Universal Robots URScript: test.script

def test():
  global _hidden_verificationVariable=0
  step_count_363709d2_59a1_48ba_b260_6a0887d41453 = 0.0
  thread Step_Counter_Thread_5b3f90a0_63de_4def_b0b2_14eef1768a44():
    while (True):
      step_count_363709d2_59a1_48ba_b260_6a0887d41453 = step_count_363709d2_59a1_48ba_b260_6a0887d41453 + 1.0
      sync()
    end
  end
  run Step_Counter_Thread_5b3f90a0_63de_4def_b0b2_14eef1768a44()
  set_gravity([0.0, 0.0, 9.82])
  motion_version_set(1)
  tool_wrench_limit_disable()
  set_tcp(p[0.0,0.0,0.161,3.1415,0.0,0.0])
  set_safety_mode_transition_hardness(1)
  set_standard_analog_input_domain(0, 1)
  set_standard_analog_input_domain(1, 1)
  set_tool_analog_input_domain(0, 1)
  set_tool_analog_input_domain(1, 1)
  set_analog_outputdomain(0, 1)
  set_analog_outputdomain(1, 1)
  set_input_actions_to_default()
  set_standard_digital_input_action(0, "freedrive")
  set_gp_boolean_input_action(0, "freedrive")
  set_runstate_standard_digital_outputs([0])
  set_runstate_configurable_digital_outputs([5])
  set_runstate_standard_digital_output_to_value(0, 1)
  set_runstate_configurable_digital_output_to_value(5, 1)
  set_runstate_configurable_digital_output_to_value(6, 2)
  set_runstate_configurable_digital_output_to_value(7, 2)
  modbus_add_signal("192.168.12.20", 255, 3, 2, "MiR_Mode", False)
  modbus_set_signal_update_frequency("MiR_Mode", 10)
  modbus_add_signal("192.168.12.20", 255, 4, 2, "MiR_State", False)
  modbus_set_signal_update_frequency("MiR_State", 10)
  modbus_add_signal("192.168.12.20", 255, 5, 2, "MiR_Error_ID", False)
  modbus_set_signal_update_frequency("MiR_Error_ID", 10)
  modbus_add_signal("192.168.12.20", 255, 7, 2, "MiR_Battery_Lvl", False)
  modbus_set_signal_update_frequency("MiR_Battery_Lvl", 10)
  modbus_add_signal("192.168.12.20", 255, 18, 2, "MiR_Mis_Queue", False)
  modbus_set_signal_update_frequency("MiR_Mis_Queue", 10)
  modbus_add_signal("192.168.12.20", 255, 1, 1, "MiR_CMD_Stop", False)
  modbus_set_signal_update_frequency("MiR_CMD_Stop", 10)
  modbus_add_signal("192.168.12.20", 255, 2, 1, "MiR_CMD_Abort", False)
  modbus_set_signal_update_frequency("MiR_CMD_Abort", 10)
  modbus_add_signal("192.168.12.20", 255, 3, 1, "MiR_CMD_Clear_Q", False)
  modbus_set_signal_update_frequency("MiR_CMD_Clear_Q", 10)
  modbus_add_signal("192.168.12.20", 255, 4, 1, "MiR_CMD_Clear_E", False)
  modbus_set_signal_update_frequency("MiR_CMD_Clear_E", 10)
  modbus_add_signal("192.168.12.20", 255, 5, 1, "MiR_CMD_Start", False)
  modbus_set_signal_update_frequency("MiR_CMD_Start", 10)
  modbus_add_signal("192.168.12.20", 255, 1001, 2, "T2O_Current_Pos", False)
  modbus_set_signal_update_frequency("T2O_Current_Pos", 10)
  modbus_add_signal("192.168.12.20", 255, 1003, 2, "T2O_Warning_ID", False)
  modbus_set_signal_update_frequency("T2O_Warning_ID", 10)
  modbus_add_signal("192.168.12.20", 255, 1005, 2, "T2O_Error_ID", False)
  modbus_set_signal_update_frequency("T2O_Error_ID", 10)
  modbus_add_signal("192.168.12.20", 255, 1019, 3, "O2T_Target_Pos", False)
  modbus_set_signal_update_frequency("O2T_Target_Pos", 10)
  modbus_add_signal("192.168.12.20", 255, 1017, 3, "O2T_Action", False)
  modbus_set_signal_update_frequency("O2T_Action", 10)
  modbus_add_signal("192.168.12.20", 255, 1000, 1, "O2T_Mis_Charge", False)
  modbus_set_signal_update_frequency("O2T_Mis_Charge", 1)
  modbus_add_signal("192.168.12.20", 255, 1004, 1, "O2T_Mis_Main", False)
  modbus_set_signal_update_frequency("O2T_Mis_Main", 1)
  modbus_add_signal("192.168.12.20", 255, 1007, 2, "T2O_Nav_Attemps", False)
  modbus_set_signal_update_frequency("T2O_Nav_Attemps", 10)
  modbus_add_signal("192.168.12.20", 255, 1009, 2, "T2O_Done", False)
  modbus_set_signal_update_frequency("T2O_Done", 10)
  modbus_add_signal("192.168.12.20", 255, 1021, 3, "O2T_Acknowledge", False)
  modbus_set_signal_update_frequency("O2T_Acknowledge", 10)
  modbus_add_signal("192.168.12.20", 255, 1011, 2, "T2O_Charging", False)
  modbus_set_signal_update_frequency("T2O_Charging", 10)
  modbus_add_signal("192.168.12.20", 255, 12, 2, "MiR_Position_X1", False)
  modbus_set_signal_update_frequency("MiR_Position_X1", 10)
  modbus_add_signal("192.168.12.20", 255, 13, 2, "MiR_Position_X2", False)
  modbus_set_signal_update_frequency("MiR_Position_X2", 10)
  modbus_add_signal("192.168.12.20", 255, 14, 2, "MiR_Position_Y1", False)
  modbus_set_signal_update_frequency("MiR_Position_Y1", 10)
  modbus_add_signal("192.168.12.20", 255, 15, 2, "MiR_Position_Y2", False)
  modbus_set_signal_update_frequency("MiR_Position_Y2", 10)
  modbus_add_signal("192.168.12.20", 255, 1023, 3, "O2T_Footprint", False)
  modbus_set_signal_update_frequency("O2T_Footprint", 10)
  modbus_add_signal("192.168.12.20", 255, 1025, 3, "O2T_ProtectOff", False)
  modbus_set_signal_update_frequency("O2T_ProtectOff", 10)
  modbus_add_signal("192.168.12.20", 255, 1027, 3, "O2T_Dock", False)
  modbus_set_signal_update_frequency("O2T_Dock", 10)
  modbus_add_signal("192.168.12.20", 255, 16, 2, "MiR_Theta_1", False)
  modbus_set_signal_update_frequency("MiR_Theta_1", 10)
  modbus_add_signal("192.168.12.20", 255, 17, 2, "MiR_Theta_2", False)
  modbus_set_signal_update_frequency("MiR_Theta_2", 10)
  modbus_add_signal("192.168.12.197", 255, 0, 0, "WM_Sensor1", False)
  modbus_set_signal_update_frequency("WM_Sensor1", 2)
  modbus_add_signal("192.168.12.197", 255, 1, 0, "WM_Sensor2", False)
  modbus_set_signal_update_frequency("WM_Sensor2", 2)
  modbus_add_signal("192.168.12.197", 255, 2, 0, "WM_Sensor3", False)
  modbus_set_signal_update_frequency("WM_Sensor3", 2)
  modbus_set_runstate_dependent_choice("MiR_CMD_Stop",0)
  modbus_set_runstate_dependent_choice("MiR_CMD_Abort",0)
  modbus_set_runstate_dependent_choice("MiR_CMD_Clear_Q",0)
  modbus_set_runstate_dependent_choice("MiR_CMD_Clear_E",0)
  modbus_set_runstate_dependent_choice("MiR_CMD_Start",0)
  modbus_set_runstate_dependent_choice("O2T_Target_Pos",0)
  modbus_set_runstate_dependent_choice("O2T_Action",0)
  modbus_set_runstate_dependent_choice("O2T_Mis_Charge",0)
  modbus_set_runstate_dependent_choice("O2T_Mis_Main",0)
  modbus_set_runstate_dependent_choice("O2T_Acknowledge",0)
  modbus_set_runstate_dependent_choice("O2T_Footprint",0)
  modbus_set_runstate_dependent_choice("O2T_ProtectOff",0)
  modbus_set_runstate_dependent_choice("O2T_Dock",0)
  set_target_payload(1.480000, [-0.002000, 0.016000, 0.051000], [0.002959, 0.002959, 0.002959, 0.000000, 0.000000, 0.000000])
  set_tool_communication(True, 115200, 0, 1, 1.5, 3.5)
  set_tool_output_mode(0)
  set_tool_digital_output_mode(0, 1)
  set_tool_digital_output_mode(1, 1)
  set_tool_voltage(24)
  global AMR_AtTarget=False
  global ARM_Referenced=False
  global PROCESS_Info=""
  global AMR_Step=0
  global STATE=4
  global AMR_Free=False
  global AMR_PosTarget=0
  global PSE_G_H=p[0, 0, 0, 0, 0, 0]
  global PSE_T=p[0.00001, -0.4, 0.30003, -0.00005, 0.00001, 0.00002]
  global PSE_R=p[0, 0, 0, 0, 0, 0]
  global AMR_PosActual=7
  global PSE_G=p[0, 0, 0, 0, 0, 0]
  global PSE_A=p[0, 0, 0, 0, 0, 0]
  global PSE_C_S=p[0, 0, 0, 0, 0, 0]
  global PSE_C_H=p[0, 0, 0, 0, 0, 0]
  global PSE_C_E=p[0, 0, 0, 0, 0, 0]
  global PSE_T_H=p[0, 0, 0, 0, 0, 0]
  global AMR_Done=True
  global STATE_Info="Idle"
  global PROCESS_Step=0
  global PSE_A_H=p[0, 0, 0, 0, 0, 0]
  global PSE_R_H=p[0, 0, 0, 0, 0, 0]
  global JNT_A=[0, 0, 0, 0, 0, 0]
  global JNT_S=[0, 0, 0, 0, 0, 0]
  global ITM_ID=0
  global JIG=0
  global JIG_Slot=0
  global OBJ_Type=0
  global PSE_Z=p[0, 0, 0, 0, 0, 0]
  global CAM_LM_Detected=True
  global CAM_LM_ID=0
  global CAM_LM_Refinmnt=False
  global CAM_Captures=0
  global CAM_Done=True
  global CAM_LM_Refined=False
  global CAM_PRM_Retries=15
  global AMR_Battery=100
  global WRK_Done=False
  global ITM_Prepared=False
  global ITM_Manipulated=False
  global AMR_Charging=False
  global Action=0
  global Task_info=""
  global Action_Info=""
  global OBJ_Picked=False
  global TM_St_Stopping="0/2/50/2"
  global STATE_Times=[37070.92578, 339840.90625, 1824.11072, 1448747.625, 26510.78125, 599104.5625, 7693.4209, 27714.24023, 201.30833, 28483.10742, 31.506, 0.258, 385.68799, 0.256, 0, 0, 0]
  global TM_St_Stopped="3/22/24/0"
  global TM_St_Resetting="0/0/30/24"
  global TM_St_Idle="16/18/25/47"
  global TM_St_Starting="0/7/21/50"
  global TM_St_Execute="6/22/25/4"
  global TM_St_Holding="0/0/3/21"
  global TM_St_Held="0/7/54/43"
  global TM_St_Unholding="0/0/0/31"
  global TM_St_Suspendin="0/0/0/0"
  global TM_St_Suspended="0/0/6/25"
  global TM_St_Unsuspend="0/0/0/0"
  global TM_St_Completin="0/2/8/13"
  global TM_St_Complete="0/7/41/54"
  global TM_St_Aborting="00/00/00/00"
  global TM_St_Aborted="00/00/00/00"
  global TM_St_Clearing="00/00/00/00"
  global CMD_Stop=False
  global STP_Info=""
  global WRK_Step=0
  global WRK_Info=""
  global AMR_FootprintID=1
  global JNT_Z=[0, 0, 0, 0, 0, 0]
  global CAM_LM_Offset=p[0, 0, 0, 0, 0, 0]
  global CAM_LM_Deviatn=p[0, 0, 0, 0, 0, 0]
  global ITM_ID_List=[1, 2, 3, 4, 5, 6, 7, 8, 9]
  global JNT_Q=[0, 0, 0, 0, 0, 0]
  global OBJ_TCP=p[0, 0.08604, 0.29117, 0, -3.14159, 0]
  global OBJ_GRP_Offset=p[0, 0, 0.15, 0, 0, 0]
  global Task_ID=0
  global PRC_Force_Decap=False
  global PRC_Reset=True
  global CAM_CNT_Obj=0
  global OBJ_Nbr=0
  global GRP_Offset=p[0, 0, 0, 0, 0, 0]
  global GRP_Open_Pos=6
  global CMD_Hold=False
  global CAM_OBJ_Color="135639"
  global JIG_Offset=p[0, 0, 0, 0, 0, 0]
  global PRM_TO_Read_BC=5
  global OBJ_Brc_OK=True
  global SERVER_IP="192.168.12.139"
  global SERVER_PORT=3002
  global POTS_IP="192.168.12.102"
  global POTS_PORT=80
  global CAM_LM_SSRack=p[0.0,0.0,0.0,0.0,0.0,0.0]
  global Cont_A_TCP=p[-0.01446224178958122,-0.6317070151410098,0.23000037816712549,-1.0906492400659007,1.4047772946314183,-1.4136947877620298]
  global Cont_B_TCP=p[0.1998,-0.5012300000000001,0.21554327201208615,-1.2092122839110917,1.2091442884557517,-1.2093098736837602]
  global Cont_C_TCP=p[0.20899409891862653,-0.36521718091627275,0.22999234057600015,-1.2337601399754432,1.1952721569824734,-1.2073910748355074]
  global Decap_TCP_align=p[-0.041471808940011026,-0.3381541550735332,0.26582523339977177,-0.8796833786644639,1.6463420679311218,-1.709080917063812]
  global FRM_Cap_SSRack=p[0.5539194080315334,0.31767425178306713,0.33208398177541654,4.365192798093082E-5,-2.191282886828362E-5,0.8765357336623923]
  global FRM_Capture_Cen=p[-0.350002433865069,0.09999194422544704,0.39999652960929194,0.27390617458472216,0.27390634457500074,1.5534190527760867]
  global FRM_Capture_IN=p[0.14713742172916425,-0.4519990092180261,0.4999842175595519,1.716719843449274E-5,-5.967839199117233E-5,-3.141512274892885]
  global FRM_Centrifuge=p[-0.7614196357228254,0.13174165134832883,-0.40322998589848,0.051405105423226086,-0.012254257775454075,1.5210337802987177]
  global FRM_Container=p[-0.5003348223692186,0.35061804815168285,0.41579001388808423,-5.092943187272062E-5,1.0145185065363121E-4,-2.764319258713288]
  global FRM_Container_b=p[-0.5003368531143569,0.35061894438330765,0.41578806736276164,-8.54682865507139E-5,1.0209605772896093E-4,-2.8884715402158117]
  global FRM_PoTS=p[-0.5403054403210852,-0.10910773999775857,0.4828,3.058497512721046E-6,2.3454853329357316E-5,-2.208510541952706]
  global FRM_Reference=p[0.0,0.0,0.0,0.0,5.936340598853489E-5,0.0]
  global FRM_SS_SSTable=p[0.20318441097787696,-0.4018484849551291,0.0986494053372641,3.321622010808724E-5,1.2630310370280906E-5,2.9057826587464487E-5]
  global FRM_SWAB=p[-0.5425658438438228,0.050215382883637555,0.4828117991467299,1.2014498510989115E-5,1.8611655946156755E-5,-2.2084947047695405]
  global FRM_weigh_scale=p[-0.3804866881697204,0.025744252835212,0.4723487455232425,-1.0445769542396123E-4,-1.924788411074358E-5,-2.1691978730572363]
  global Home_Center=p[8.153119343667444E-6,-0.39999432384352546,0.2999959692487133,2.5646064776662724E-5,4.3940218780729606E-7,1.0264337438974612E-5]
  global Position1=p[-0.013283381383284571,-0.5604926192866768,0.38388715699602394,4.2328981461085945E-5,2.7078270325215812E-5,-3.7205146207707955E-5]
  global Position2=p[0.20351564705697425,-0.4203376101670667,0.3838762041571461,3.798288302544451E-5,4.704460451857417E-5,4.231147149799096E-6]
  global Position3=p[0.20350843333470736,-0.29021893349684563,0.38387753498709576,1.6019315164720892E-6,5.362200339537394E-5,1.3194338684148116E-5]
  global SAF_ULM_Back=p[0.0,0.25,0.0,-1.5707963267948966,0.0,0.0]
  global SAF_ULM_Bottom=p[0.0,0.0,0.175,0.0,-3.1411853059779946,6.144646783253781E-5]
  global SAF_ULM_Front=p[0.0,-0.8,0.0,1.5707963267948966,0.0,0.0]
  global SAF_ULM_Left=p[0.4,0.0,0.0,0.0,1.5707963267948966,0.0]
  global SAF_ULM_Right=p[-0.4,0.0,0.0,0.0,-1.5707963267948966,0.0]
  global Swab_Hol_NewApp=p[0.24367285099070987,-0.39538254967913455,0.1791890228280021,9.694511507909782E-6,-1.918651308171816E-5,-8.936699871509937E-5]
  global Swab_Holder=p[0.24295783117309838,-0.3013564682530984,0.1852322720229175,2.781519887568103E-5,4.9787017742599154E-5,-4.37903285531786E-5]
  global Swab_Holder_App=p[0.2429619714479549,-0.37982819606840945,0.18525382710668278,1.9222871262119376E-5,1.6223417670491008E-5,-5.4734062838048446E-5]
  global Swab_New_FlipAp=p[0.2397112683246373,-0.4131931547204771,0.1791901367353106,-3.2195134883720305E-6,5.5826332611522435E-5,3.121155597546625]
  global Swab_New_FlipHL=p[0.24201994270482732,-0.3016396679914842,0.1792041435801504,-5.840580747813655E-5,7.149594627182296E-5,3.1212173415187716]
  global Swab_flip_app=p[0.2429388733172488,-0.30137068448833126,0.2604132558601291,2.6401756342031075E-4,-5.484374510519208E-5,3.1254804120366084]
  global Swab_flip_hold=p[0.24294214110481466,-0.30136164018491357,0.18562266741928893,2.522236506414148E-4,-7.112060556159522E-5,3.1255321079816243]
  global Swab_holder_New=p[0.24365536646762584,-0.2997701233168029,0.17918094816818864,3.214234787213423E-5,4.175157661863989E-5,-5.646064180042735E-5]
  global Swab_take=p[0.06323186369735694,-0.63186492852859,0.1186768659332022,-0.0941457732311389,0.09836792894816203,-1.517326737506051]
  global Swab_take_appro=p[0.06320391400111934,-0.6318588436631464,0.19565149002631285,-0.09417297851843164,0.09839511960035544,-1.5173200644593776]
  global Trigger=p[0.0,0.0,0.0,0.0,0.0,0.0]
  global ULM_3FG=p[-0.030765235416747628,-0.34863465891472667,0.113,7.284395488044268E-6,3.273453749838684E-5,-1.4353257859996407]
  global ULM_Cap_Bin=p[-0.09250864937066318,-0.4278810928466919,0.11,0.012411963638116327,0.0011373915061224443,2.7934337459497622]
  global ULM_Cent_Racks=p[-0.18545280836253272,-0.6127182427471424,0.0092,-2.5489681018192384E-4,1.5011949774034494E-5,0.002017828229688311]
  global ULM_Input=p[0.24211961776286645,-0.49122804302630946,0.069,-0.0024427818584600467,0.009435707692609437,1.553764323389261]
  global ULM_NoK=p[-0.13173558762545426,-0.4223773499069831,0.1783860505865236,-0.013295546620598609,-0.0036702711105456223,-3.139406935149283]
  global ULM_Output=p[-0.03848915736486644,-0.4320501686344275,0.0,-6.433221303631731E-5,4.4743073056790854E-4,-3.1218466433891914]
  global ULM_SS_Jig=p[0.20042235181396445,-0.401422571467659,0.10172961048670293,-0.004383916608756479,-0.025399236865877438,0.14513627174952076]
  global swab_brk1=p[-0.038192766284940796,-0.35032292650225555,0.1065863357332553,-1.0289939058230132E-4,2.813749403516853,1.8382182448234926E-4]
  global uLM_Cap_SSRack=p[0.20881778585250285,-0.4048217020440386,0.5540171693698591,2.8523205665698764E-5,1.4454354491120644E-5,-0.034379521481452686]
  global uLM_SS_PickPlc=p[0.16950832747543634,-0.42825836359263725,0.10175705391961387,4.604858547296167E-4,-6.723821859499963E-4,-2.834490280150995]
  # begin: URCap Installation Node
  #   Source: UR Connect, 2.3.3, Universal Robots
  #   Type: UR Connect
  myurRPC = rpc_factory("xmlrpc","http://127.0.0.1:40474")
  # end: URCap Installation Node
  # begin: URCap Installation Node
  #   Source: Robotiq_Grippers, 3.17.0.105337, Robotiq Inc.
  #   Type: Vacuum
  #################################################
  # Vacuum Grip Check
  #################################################

  vacuumGripCheckThread1 = 0
  vacuumGripCheckThread2 = 0
  vacuumGripCheckThread3 = 0
  vacuumGripCheckThread4 = 0
  vacuumGripCheckThread1Running = False
  vacuumGripCheckThread2Running = False
  vacuumGripCheckThread3Running = False
  vacuumGripCheckThread4Running = False
  vacuumGripCheckSocketId = "1"
  vacuumGripCheckThreadStarted = False

  thread vacuumGripCheck():
    gripper_socket = vacuumGripCheckSocketId
    vacuumGripCheckThreadStarted = True

    while (True):
      objectDetectedDebounceCtr = 0

      while (objectDetectedDebounceCtr < 3):
        if(rq_is_vacuum_obj_detected(gripper_socket="1")):
          objectDetectedDebounceCtr = objectDetectedDebounceCtr + 1
        else:
          objectDetectedDebounceCtr = 0
        end
        sleep(0.1)
      end

      objectNotDetectedDebounceCtr = 0

      while objectNotDetectedDebounceCtr < 3:
        if (not rq_is_vacuum_obj_detected(gripper_socket="1")):
          objectNotDetectedDebounceCtr = objectNotDetectedDebounceCtr + 1
        else:
          objectNotDetectedDebounceCtr = 0
        end
        sleep(0.1)
      end

      socket_open("127.0.0.1",29999,"dashboardServerSocket")
      socket_send_line("pause","dashboardServerSocket")
      socket_send_string("popup Vacuum grip check has detected an object drop.", "dashboardServerSocket")
      socket_send_byte(10, "dashboardServerSocket")
      socket_close("dashboardServerSocket")

      sleep(0.008)
    end
  end

  def startVacuumGripCheckThread(gripperId="1"):
    vacuumGripCheckSocketId = gripperId
    threadHandle = run vacuumGripCheck()
    waitForVacuumGripCheckThreadStarted()
    return threadHandle
  end

  def stopVacuumGripCheckThread(threadHandle):
    kill threadHandle
  end

  def waitForVacuumGripCheckThreadStarted():
    while (not(vacuumGripCheckThreadStarted)):
      sleep(0.008)
    end
    vacuumGripCheckThreadStarted = False
  end
  #################################################
  # End - Vacuum Grip Check
  #################################################

  #################################################
  # Stops the pump on a distance travelled
  #################################################
  global stopPumpDistance = 100
  global stopPumpSocketId = "0"
  global stopPumpThreadStarted = [False, False, False, False]
  global stopPumpThreadHandles = [0, 0, 0, 0]

  thread stopPumpOnDistanceTravelled():
    distance = stopPumpDistance
    socketId = stopPumpSocketId
    stopPumpThreadStarted[rq_socket_to_index(socketId)] = True

    measuredDistance = waitForDistanceTravelled(distance)

    rq_stop(socketId)

    stopPumpThreadStarted[rq_socket_to_index(socketId)] = False
  end

  def waitForDistanceTravelled(distance):
    startingPose = get_actual_tcp_pose()
    measuredDistance = 0
    while (measuredDistance < distance):
      sleep(0.1)
      measuredDistance = point_dist(get_actual_tcp_pose(), startingPose)
    end

    return measuredDistance
  end

  def startStopPumpOnDistanceTravelledThread(distance, gripper_socket="1"):
    if (stopPumpThreadStarted[rq_socket_to_index(gripper_socket)]):
      return 0
    end

    global stopPumpDistance = distance
    global stopPumpSocketId = gripper_socket
    stopPumpThreadHandles[rq_socket_to_index(gripper_socket)] = run stopPumpOnDistanceTravelled()
    waitForStopPumpOnDistanceTravelledThreadStarted(gripper_socket)
    return stopPumpThreadHandles[rq_socket_to_index(gripper_socket)]
  end

  def waitForStopPumpOnDistanceTravelledThreadStarted(gripper_socket="1"):
    while (not(stopPumpThreadStarted[rq_socket_to_index(gripper_socket)])):
      sleep(0.008)
    end
  end

  def stopStopPumpOnDistanceTravelledThread(gripper_socket="1"):
    handle = stopPumpThreadHandles[rq_socket_to_index(gripper_socket)]
    threadIsRunning = stopPumpThreadStarted[rq_socket_to_index(gripper_socket)]
    if (threadIsRunning):
      kill handle
      clear_socket_buffer(gripper_socket, 0.01)
      stopPumpThreadHandles[rq_socket_to_index(gripper_socket)] = 0
    end
  end
  #################################################
  # End - Stops the pump on a distance travelled
  #################################################

  #################################################
  # Vacuum general functions
  #################################################
  def rq_wait_for_vacuum_object_detected(gripper_socket="1"):
      while (not rq_is_vacuum_obj_detected(gripper_socket)):
          if (rq_is_vacuum_timeout(gripper_socket)):
              return False
          end
          sleep(0.008)
      end
      return True
  end

  def rq_wait_for_vacuum_object_secured(gripper_socket="1"):
      while (not rq_is_vacuum_obj_secured(gripper_socket)):
          if (rq_is_vacuum_timeout(gripper_socket)):
              return False
          end
          sleep(0.008)
      end
      return True
  end

  def rq_wait_for_vacuum_object_suction_complete(gripper_socket="1"):
      remaining_retries = 50

       # Wait for suction started
      while (not rq_is_vacuum_obj_in_suction(gripper_socket) and
             not rq_is_vacuum_obj_detected(gripper_socket) and
             remaining_retries > 0):
          sleep(0.01)
          remaining_retries = remaining_retries - 1
      end

      # Wait for suction completed
      while (rq_is_vacuum_obj_in_suction(gripper_socket)):
          if (rq_is_vacuum_timeout(gripper_socket)):
              return False
          end
          sleep(0.01)
      end

      return True
  end

  def rq_wait_for_vacuum_object_not_detected(gripper_socket="1"):
      while (rq_is_vacuum_obj_detected(gripper_socket)):
          sleep(0.01)
      end
  end

  def rq_is_vacuum_obj_detected(gripper_socket="1"):
      gOBJ = rq_get_var("OBJ", 1, gripper_socket)
      sleep(0.008)
      return is_vacuum_OBJ_object_detected(gOBJ)
  end

  def rq_is_vacuum_obj_secured(gripper_socket="1"):
      gOBJ = rq_get_var("OBJ", 1, gripper_socket)
      sleep(0.008)
      return is_vacuum_OBJ_object_secured(gOBJ)
  end

  def rq_is_vacuum_obj_in_suction(gripper_socket="1"):
      gOBJ = rq_get_var("OBJ", 1, gripper_socket)
      sleep(0.008)

      if(is_vacuum_OBJ_object_in_motion(gOBJ)):
          return True
      else:
          return False
      end
  end

  def rq_is_vacuum_timeout(gripper_socket="1"):
      gFLT = rq_get_var("FLT", 2, gripper_socket)
      sleep(0.008)

      if(gFLT ==6):
          return True
      end

      return False
  end

  def is_vacuum_OBJ_object_in_motion(gOBJ):
      if (gOBJ == 0):
          return True
      end

      return False
  end

  def is_vacuum_OBJ_object_detected(gOBJ):
      if (gOBJ == 1 or gOBJ == 2):
          return True
      end

      return False
  end

  def is_vacuum_OBJ_object_secured(gOBJ):
      if (gOBJ == 2):
          return True
      end

      return False
  end

  def rq_set_pressure_timeout_minimum_vacuum(pressure, timeout, minimum, gripper_socket="1"):
      rq_set_pos_spd_for(pressure, timeout, minimum, gripper_socket)
  end

  def rq_set_vacuum_and_wait(pressure, timeout, minimum, mode, gripper_socket="1"):
      rq_set_pressure_timeout_minimum_vacuum(pressure, timeout, minimum, gripper_socket)
      gPRE = rq_get_var("PRE", 3, gripper_socket)
      while (gPRE != pressure):
          rq_set_pressure_timeout_minimum_vacuum(pressure, timeout, minimum, gripper_socket)
          sleep(0.008)
          gPRE = rq_get_var("PRE", 3, gripper_socket)
      end

      rq_set_gripper_mode(mode, gripper_socket)
      gMOD = rq_get_var("MOD", 3, gripper_socket)
      while (gMOD != mode):
          rq_set_gripper_mode(mode, gripper_socket)
          sleep(0.008)
          gMOD = rq_get_var("MOD", 3, gripper_socket)
     end
  end

  def is_FLT_vacuum_timeout(gFLT):
    if (gFLT == 6):
        return True
    end

    return False
  end

  def is_continuous_grip(maximum_vacuum):
    return maximum_vacuum == 0
  end

  def rq_vacuum_release(advanced_mode=False, shutoff_distance_cm=5, wait_for_object_released=True, gripper_socket="1"):
    local shutoff_distance = scale(shutoff_distance_cm, [0, 99], [0.00, 0.99])
    local pressure = 255
    local minimum = 0
    local timeout = 255
    rq_vacuum_release_raw(advanced_mode, pressure, minimum, timeout, shutoff_distance, wait_for_object_released, gripper_socket)
  end

  def rq_vacuum_release_raw(advanced_mode, pressure, minimum, timeout, shutoff_distance, wait_for_object_released, gripper_socket):
    rq_reset_fault_and_activate(gripper_socket)

    if advanced_mode:
      rq_set_vacuum_and_wait(pressure, timeout, minimum, 1, gripper_socket)
    else:
      rq_set_vacuum_and_wait(pressure, timeout, minimum, 0, gripper_socket)
    end

    # The following patch is for Robotiq's Camera issue when communication is lost, but not the activation
    # the communication driver reset the GTO bit
    rq_set_GTO_and_wait(1, gripper_socket)

    if wait_for_object_released:
      while (rq_is_vacuum_obj_detected(gripper_socket)):

        if advanced_mode:
          rq_set_vacuum_and_wait(pressure, timeout, minimum, 1, gripper_socket)
        else:
          rq_set_vacuum_and_wait(pressure, timeout, minimum, 0, gripper_socket)
        end

        # The following patch is for Robotiq's Camera issue when communication is lost, but not the activation
        # the communication driver reset the GTO bit
        rq_set_GTO_and_wait(1, gripper_socket)
        sleep(0.01)
      end
    end

    if advanced_mode:
      startStopPumpOnDistanceTravelledThread(shutoff_distance, gripper_socket)
    end
  end

  def rq_vacuum_grip(advanced_mode=False, maximum_vacuum=60, minimum_vacuum=40, timeout_ms=3000, wait_for_object_detected=True, gripper_socket="1"):
    local pressure = scale(maximum_vacuum, [0, 100], [100, 0])
    local minimum = scale(minimum_vacuum, [0, 100], [100, 0])
    local timeout = scale(timeout_ms, [0, 25500], [0, 255])
    rq_vacuum_grip_raw(advanced_mode, pressure, minimum, timeout, gripper_socket)
    if wait_for_object_detected:
          suction_completed = rq_wait_for_vacuum_object_suction_complete(gripper_socket)
          if(not suction_completed):
              rq_set_var("GTO", 0, gripper_socket)
          end
    end
  end

  def rq_vacuum_grip_raw(advanced_mode, pressure, minimum, timeout, gripper_socket):
    stopStopPumpOnDistanceTravelledThread(gripper_socket)
    rq_reset_fault_and_activate(gripper_socket)

    if advanced_mode:
      rq_set_vacuum_and_wait(pressure, timeout, minimum, 1, gripper_socket)
    else:
      rq_set_vacuum_and_wait(pressure, timeout, minimum, 0, gripper_socket)
    end

    rq_set_GTO_and_wait(1, gripper_socket)
  end

  def rq_reset_fault_and_activate(gripper_socket):
      gFLT = rq_get_var("FLT", 2, gripper_socket)

      if(not is_FLT_no_fault(gFLT)):
          if(is_FLT_vacuum_timeout(gFLT)):
              rq_set_GTO_and_wait(0, gripper_socket)
          elif(is_FLT_faulted(gFLT)):
              rq_set_GTO_and_wait(0, gripper_socket)
              rq_set_var("ACT", 1, gripper_socket)
          end
      elif(not rq_is_gripper_activated(gripper_socket)):
          rq_set_GTO_and_wait(0, gripper_socket)
          rq_set_var("ACT", 1, gripper_socket)
      end
  end
  #################################################
  # End - Vacuum general functions
  #################################################
  vacuumGripCheckWarningTitle = "Vacuum grip check"
  vacuumGripCheckWarningMessage = "Vacuum gripper object lost"
  vacuumGripTimeoutTitle = "Vacuum gripper fault"
  vacuumGripTimeoutMessage = "Grip has timed out"
  # end: URCap Installation Node
  # begin: URCap Installation Node
  #   Source: SensoPart VISOR Robotic, 2.0.6, SensoPart Industriesensorik GmbH
  #   Type: VISOR Robotic
  visor_xml_rpc_client = rpc_factory("xmlrpc", "http://127.0.0.1:" + to_str(42023) + "/RPC2\")

  #######################################
  # Settings
  visor__errInterrupt = True
  visor__debugLvl = 1

  #######################################
  # Variables
  visor__varSendReqOk = [False,False,False,False,False,False,False,False]
  visor__varRespOk = [False,False,False,False,False,False,False,False]
  visor__partsFound = [0,0,0,0,0,0,0,0]
  visor__objPos_1 = [ p[0,0,0,0,0,0], p[0,0,0,0,0,0], p[0,0,0,0,0,0], p[0,0,0,0,0,0], p[0,0,0,0,0,0], p[0,0,0,0,0,0], p[0,0,0,0,0,0], p[0,0,0,0,0,0], p[0,0,0,0,0,0], p[0,0,0,0,0,0] ]
  visor__objPos_2 = [ p[0,0,0,0,0,0], p[0,0,0,0,0,0], p[0,0,0,0,0,0], p[0,0,0,0,0,0], p[0,0,0,0,0,0], p[0,0,0,0,0,0], p[0,0,0,0,0,0], p[0,0,0,0,0,0], p[0,0,0,0,0,0], p[0,0,0,0,0,0] ]
  visor__objPos_3 = [ p[0,0,0,0,0,0], p[0,0,0,0,0,0], p[0,0,0,0,0,0], p[0,0,0,0,0,0], p[0,0,0,0,0,0], p[0,0,0,0,0,0], p[0,0,0,0,0,0], p[0,0,0,0,0,0], p[0,0,0,0,0,0], p[0,0,0,0,0,0] ]
  visor__objPos_4 = [ p[0,0,0,0,0,0], p[0,0,0,0,0,0], p[0,0,0,0,0,0], p[0,0,0,0,0,0], p[0,0,0,0,0,0], p[0,0,0,0,0,0], p[0,0,0,0,0,0], p[0,0,0,0,0,0], p[0,0,0,0,0,0], p[0,0,0,0,0,0] ]
  visor__objPos_5 = [ p[0,0,0,0,0,0], p[0,0,0,0,0,0], p[0,0,0,0,0,0], p[0,0,0,0,0,0], p[0,0,0,0,0,0], p[0,0,0,0,0,0], p[0,0,0,0,0,0], p[0,0,0,0,0,0], p[0,0,0,0,0,0], p[0,0,0,0,0,0] ]
  visor__objPos_6 = [ p[0,0,0,0,0,0], p[0,0,0,0,0,0], p[0,0,0,0,0,0], p[0,0,0,0,0,0], p[0,0,0,0,0,0], p[0,0,0,0,0,0], p[0,0,0,0,0,0], p[0,0,0,0,0,0], p[0,0,0,0,0,0], p[0,0,0,0,0,0] ]
  visor__objPos_7 = [ p[0,0,0,0,0,0], p[0,0,0,0,0,0], p[0,0,0,0,0,0], p[0,0,0,0,0,0], p[0,0,0,0,0,0], p[0,0,0,0,0,0], p[0,0,0,0,0,0], p[0,0,0,0,0,0], p[0,0,0,0,0,0], p[0,0,0,0,0,0] ]
  visor__objPos_8 = [ p[0,0,0,0,0,0], p[0,0,0,0,0,0], p[0,0,0,0,0,0], p[0,0,0,0,0,0], p[0,0,0,0,0,0], p[0,0,0,0,0,0], p[0,0,0,0,0,0], p[0,0,0,0,0,0], p[0,0,0,0,0,0], p[0,0,0,0,0,0] ]
  visor__easyPickNodeId = ""
  visor__easyPickDeviceId = 0

  #######################################
  # Public functions
  def visor_isSendReqOk(device_id):
    visor__checkDeviceId(device_id)
    return visor__varSendReqOk[device_id - 1]
  end

  def visor_isResponseOk(device_id):
    visor__checkDeviceId(device_id)
    return visor__varRespOk[device_id - 1]
  end

  def visor_getResponse(device_id):
    visor__checkDeviceId(device_id)
    return visor_xml_rpc_client.Update.getResponse(device_id - 1)
  end

  def visor_terminal(device_id, request, opt_timeout = 6000):
    visor__checkDeviceId(device_id)
    while (not visor__sendRequest(device_id - 1, opt_timeout, request)):
      if visor__popup("Send terminal request failed"):
        return None
      end
    end
  end

  def visor_changeJob(device_id, jobName, opt_timeout = 6000):
    visor__checkDeviceId(device_id)
    visor__sendReqWaitSuccess(device_id - 1, opt_timeout, "CJN1" + visor__valToStr(str_len(jobName), 3) + jobName, "Send change job request failed","Change job failed")
  end

  def visor_trigger(device_id, opt_timeout = 6000, opt_setup = "fix"):
    visor__checkDeviceId(device_id)

    # Reset variables
    visor__partsFound[device_id -1] = 0

    # Execute trigger
    if (opt_setup =="arm"):
      visor__sendReqWaitSuccess(device_id - 1, opt_timeout, "TRR100" + visor__poseToVisorStr(get_actual_tcp_pose()), "Send trigger failed","Trigger not successful")
    else:
      visor__sendReqWaitSuccess(device_id - 1, opt_timeout, "TRX00", "Send trigger failed","Trigger not successful")
    end

    # Send and response ok?
    if (not (visor__varSendReqOk[device_id - 1] and visor__varRespOk[device_id - 1])):
      visor__logMsg("VISOR, send trigger failed or fail response", True)
      visor__popup("Send trigger failed or fail response<br>Perhaps the connection was interrupted or the VISOR was not ready")
      return None
    end

    # Parse trigger response
    if (not visor_xml_rpc_client.Update.parseTriggerResult(device_id - 1)):
      visor__logMsg("VISOR, unable to parse trigger result, maybe wrong format", True)
      visor__popup("Incorrect Trigger Response<br>Did you configure the telegram for the used detector in SensoConfig correctly?")
      return None
    end
    visor__partsFound[device_id - 1] = visor_xml_rpc_client.Update.getTriggerPartsFound(device_id - 1)
    local i = 0
    while (i < visor__partsFound[device_id - 1]):
      visor__setObjPos(device_id, visor_xml_rpc_client.Update.getTriggerObjPos(device_id - 1, i), i)
      i = i + 1
    end
  end

  def visor_partsFound(device_id):
    visor__checkDeviceId(device_id)
    return visor__partsFound[device_id - 1]
  end

  def visor_resetResult(device_id):
    visor__checkDeviceId(device_id)
    visor__partsFound[device_id -1] = 0
  end

  def visor_getObjPos(device_id, idx):
    visor__checkDeviceId(device_id)
    visor__checkResultIdx(idx)
    return visor__getObjPos(device_id, idx)
  end

  def visor_getPose2d(device_id, idx, opt_refPose=p[0,0,0,0,0,0]):
    visor__checkDeviceId(device_id)
    visor__checkResultIdx(idx)
    local objPos = visor__getObjPos(device_id, idx)
    local refPose = pose_trans(opt_refPose, p[0,0,0,0,0,d2r(objPos[5])])
    return p[objPos[0] / 1000, objPos[1] / 1000, refPose[2], refPose[3], refPose[4], refPose[5]]
  end

  def visor_getPose3d(device_id, idx):
    visor__checkDeviceId(device_id)
    visor__checkResultIdx(idx)
    local objPos = visor__getObjPos(device_id, idx)
    local angles = rpy2rotvec([d2r(objPos[3]), d2r(objPos[4]), d2r(objPos[5])])
    return p[objPos[0] / 1000, objPos[1] / 1000, objPos[2] / 1000, angles[0], angles[1], angles[2]]
  end

  def visor_getAdditionalData(device_id, opt_idx=999):
    visor__checkDeviceId(device_id)
    return visor_xml_rpc_client.Update.getTriggerAdditionalData(device_id - 1, opt_idx)
  end

  def visor_getCalibSetImgPose(setNo):
    return visor_xml_rpc_client.Update.getCalibSetImagePose(setNo)
  end

  def visor_easyPickUpdate(device_id, param, value):
    visor__checkDeviceId(device_id)
    return visor_xml_rpc_client.Update.setEasyPickUpdate(device_id - 1, param, to_str(value))
  end

  def visor_activateOffset(device_id, detector_no, offset_mode, opt_timeout = 6000):
    visor__checkDeviceId(device_id)

    # Check detector number
    if (detector_no < 0) or (detector_no > 999):
      visor__logMsg("VISOR, invalid detector no: " + to_str(detector_no), True)
      visor__popup("Invalid detector no")
      halt
    end

    # Check offset_mode
    if (offset_mode != 0) and (offset_mode != 3):
      visor__logMsg("VISOR, invalid offset mode: " + to_str(offset_mode), True)
      visor__popup("Invalid offset mode")
      halt
    end

    # Send request
    local spp_request = "SPP" + visor__valToStr(detector_no, 3) + "030" + "00001" + to_str(offset_mode)
    visor__sendReqWaitSuccess(device_id - 1, opt_timeout, spp_request, "Activate offset failed", "Activate offset failed")

    return visor__varRespOk[device_id - 1]
  end

  def visor_teachOffset(device_id, detector_no, offset_pose, opt_timeout = 6000):
    visor__checkDeviceId(device_id)

    # Check detector number
    if (detector_no < 0) or (detector_no > 999):
      visor__logMsg("VISOR, invalid detector no: " + to_str(detector_no), True)
      visor__popup("Invalid detector nr")
      halt
    end

    # Send request
    local spp_request = "SPP" + visor__valToStr(detector_no, 3) + "035" + "00048" + visor__poseToVisorStr(offset_pose)
    visor__sendReqWaitSuccess(device_id - 1, opt_timeout, spp_request, "Teach offset failed", "Teach offset failed")

    return visor__varRespOk[device_id - 1]
  end

  def visor_calcCenter3d(device_id, visor1_pose, visor2_pose, opt_timeout = 6000):
  	visor__checkDeviceId(device_id)

  	local rf_mf_pose = p[0,0,0,0,0,0]
  	local mid_pose = p[0,0,0,0,0,0]

  	# get rm_mf
  	visor__sendReqWaitSuccess(device_id - 1, opt_timeout, "CGP1015", "Calculate center 3D not successful" , "Calculate center 3D not successful")
      local response = visor_xml_rpc_client.Update.getResponse(device_id - 1)
      if (visor__varSendReqOk[device_id - 1] and visor__varRespOk[device_id - 1]):
        local loopIdx = 0
        while (loopIdx < 6):
          rf_mf_pose[loopIdx] = to_num(str_sub(response,18+(loopIdx*8),8))/1000
          if (loopIdx > 2) and (loopIdx < 6):
            rf_mf_pose[loopIdx] = d2r(rf_mf_pose[loopIdx])
          end
          loopIdx = loopIdx + 1
        end
      end
      local axis_angle = rpy2rotvec([(rf_mf_pose[3]),(rf_mf_pose[4]),(rf_mf_pose[5])])
  	rf_mf_pose[3] = axis_angle[0]
  	rf_mf_pose[4] = axis_angle[1]
  	rf_mf_pose[5] = axis_angle[2]

  	# invert rf_mf_pose
      local rm_mf_pose_inverse = pose_inv(rf_mf_pose)

      # transform visor poses to measurement frame
      local visor1_pose_trans = pose_trans(rm_mf_pose_inverse, visor1_pose)
      local visor2_pose_trans = pose_trans(rm_mf_pose_inverse, visor2_pose)

      # calculate angle in measurement frame
      local dx = (visor2_pose_trans[0]-visor1_pose_trans[0])
      local dy = (visor2_pose_trans[1]-visor1_pose_trans[1])
      mid_pose[5] = atan(dy/dx)
      axis_angle = rpy2rotvec([(mid_pose[3]),(mid_pose[4]),(mid_pose[5])])
      mid_pose[3] = axis_angle[0]
  	mid_pose[4] = axis_angle[1]
  	mid_pose[5] = axis_angle[2]

      # transform back to robot frame
      mid_pose = pose_trans(rf_mf_pose, mid_pose)

      # center of x, y, z
      mid_pose[0] = (visor1_pose[0]+visor2_pose[0])/2
      mid_pose[1] = (visor1_pose[1]+visor2_pose[1])/2
      mid_pose[2] = (visor1_pose[2]+visor2_pose[2])/2

  	return mid_pose
  end

  def visor_easyPickCheckIdent(node_id, device_id):
    return (visor__easyPickNodeId == node_id) and (visor__easyPickDeviceId == device_id)
  end

  def visor_easyPickSetIdent(node_id, device_id):
    visor__easyPickNodeId = node_id
    visor__easyPickDeviceId = device_id
  end

  #######################################
  # Private functions
  def visor__checkDeviceId(device_id):
    if (device_id < 1) or (device_id > 8):
      visor__logMsg("VISOR, invalid device id: " + to_str(device_id), True)
      visor__popup("Invalid device id")
      halt
    end
  end

  def visor__checkResultIdx(idx):
    if (idx < 0) or (idx > 9):
      visor__logMsg("VISOR, invalid result index: " + to_str(idx), True)
      visor__popup("Invalid result index")
      halt
    end
  end

  def visor__logMsg(message, important=False):
    if (visor__debugLvl == 2) or important:
      textmsg(message)
    end
  end

  def visor__popup(message, warn=False, err=True):
    if visor__errInterrupt:
      popup(message, title="VISOR", warning=warn, error=err, blocking=True)
    end
    return (not visor__errInterrupt)
  end

  def visor__sendReqWaitSuccess(device_id, timeout, request, msgSendErr, msgRespErr):
    while True:
      if visor__sendRequest(device_id, timeout, request):
        if visor__varRespOk[device_id]:
          return None
        else:
          if visor__popup(msgRespErr, True, False):
            return None
          end
        end
      else:
        if visor__popup(msgSendErr):
          return None
        end
      end
    end
  end

  def visor__sendRequest(device_id, timeout, request):
    visor__logMsg("VISOR, send_request: " + request)
    visor__varSendReqOk[device_id] = visor_xml_rpc_client.Update.sendRequest(device_id, timeout, request)
    visor__varRespOk[device_id] = visor_xml_rpc_client.Update.isResponseOk(device_id)
    local response = visor_xml_rpc_client.Update.getResponse(device_id)
    visor__logMsg("VISOR, response: " + response)
    return visor__varSendReqOk[device_id]
  end

  def visor__valToStr(val, digits=0):
    local s = to_str(val)
    local delta = digits - str_len(s)
    local negative = False
    if (str_at(s, 0) == "-"):
      negative = True
      s = str_sub(s, 1)
    end
    while (delta > 0):
      s = "0" + s
      delta = delta -1
    end
    if negative:
      s = "-" + s
    end
    return s
  end

  def visor__setObjPos(device_id, pose, idx):
    if (device_id == 1):
      visor__objPos_1[idx] = pose
    elif (device_id == 2):
      visor__objPos_2[idx] = pose
    elif (device_id == 3):
      visor__objPos_3[idx] = pose
    elif (device_id == 4):
      visor__objPos_4[idx] = pose
    elif (device_id == 5):
      visor__objPos_5[idx] = pose
    elif (device_id == 6):
      visor__objPos_6[idx] = pose
    elif (device_id == 7):
      visor__objPos_7[idx] = pose
    elif (device_id == 8):
      visor__objPos_8[idx] = pose
    end
  end

  def visor__getObjPos(device_id, idx):
    if (device_id == 1):
      return visor__objPos_1[idx]
    elif (device_id == 2):
      return visor__objPos_2[idx]
    elif (device_id == 3):
      return visor__objPos_3[idx]
    elif (device_id == 4):
      return visor__objPos_4[idx]
    elif (device_id == 5):
      return visor__objPos_5[idx]
    elif (device_id == 6):
      return visor__objPos_6[idx]
    elif (device_id == 7):
      return visor__objPos_7[idx]
    elif (device_id == 8):
      return visor__objPos_8[idx]
    end
  end

  def visor__poseToVisorStr(tcpPose, useAxisAngle=False):
    # Convert to RPY, default VISOR configuration
    local rpy = rotvec2rpy([tcpPose[3], tcpPose[4], tcpPose[5]])

    poseStr = ""
    i = 0
    while (i < 6):
      if (i > 2):
        # Rotation, use RPY or axis angle and multiply by 1000
        if (not useAxisAngle):
          tcpPose[i] = r2d(rpy[i-3])
        end
        tcpPose[i] = floor(tcpPose[i] * 1000)
      else:
        # Location, convert to [mm] and multiply by 1000
        tcpPose[i] = floor(tcpPose[i] * 1000000)
      end
      # Convert value to valid format (prefixing with '0')
      # and add to pose string
      poseStr = poseStr + visor__valToStr(tcpPose[i], 8)
      i = i + 1
    end
    return poseStr
  end
  # end: URCap Installation Node
  # begin: URCap Installation Node
  #   Source: Robotiq_Grippers, 3.17.0.105337, Robotiq Inc.
  #   Type: Gripper
  rq_gripper_socket_ip_address = "127.0.0.1"
  rq_gripper_socket_port = 63352

  rq_comm_check_fail_counter = [0, 0, 0, 0]

  rq_read_act = [-1, -1, -1, -1]
  rq_read_gto = [-1, -1, -1, -1]
  rq_read_for = [-1, -1, -1, -1]
  rq_read_spe = [-1, -1, -1, -1]
  rq_read_obj = [-1, -1, -1, -1]
  rq_read_sta = [-1, -1, -1, -1]
  rq_read_flt = [-1, -1, -1, -1]
  rq_read_pos = [-1, -1, -1, -1]
  rq_read_pre = [-1, -1, -1, -1]
  rq_read_lbp = [-1, -1, -1, -1]
  rq_read_lrd = [-1, -1, -1, -1]
  rq_read_lbl = [-1, -1, -1, -1]
  rq_read_lgn = [-1, -1, -1, -1]
  rq_read_msc = [-1, -1, -1, -1]
  rq_read_mod = [-1, -1, -1, -1]
  rq_read_cou = [-1, -1, -1, -1]
  rq_read_ncy = [-1, -1, -1, -1]
  rq_read_dst = [-1, -1, -1, -1]
  rq_read_pco = [-1, -1, -1, -1]

  rq_string_initial_value = "N/A"

  rq_read_snu_1 = rq_string_initial_value
  rq_read_snu_2 = rq_string_initial_value
  rq_read_snu_3 = rq_string_initial_value
  rq_read_snu_4 = rq_string_initial_value

  rq_read_fwv_1 = rq_string_initial_value
  rq_read_fwv_2 = rq_string_initial_value
  rq_read_fwv_3 = rq_string_initial_value
  rq_read_fwv_4 = rq_string_initial_value

  rq_read_ver_1 = rq_string_initial_value
  rq_read_ver_2 = rq_string_initial_value
  rq_read_ver_3 = rq_string_initial_value
  rq_read_ver_4 = rq_string_initial_value

  rq_read_act_req = [True, True, True, True]
  rq_read_gto_req = [True, True, True, True]
  rq_read_for_req = [True, True, True, True]
  rq_read_spe_req = [True, True, True, True]
  rq_read_obj_req = [True, True, True, True]
  rq_read_sta_req = [True, True, True, True]
  rq_read_flt_req = [True, True, True, True]
  rq_read_pos_req = [True, True, True, True]
  rq_read_pre_req = [True, True, True, True]
  rq_read_lbp_req = [True, True, True, True]
  rq_read_lrd_req = [True, True, True, True]
  rq_read_lbl_req = [True, True, True, True]
  rq_read_lgn_req = [True, True, True, True]
  rq_read_msc_req = [True, True, True, True]
  rq_read_mod_req = [True, True, True, True]
  rq_read_cou_req = [True, True, True, True]
  rq_read_ncy_req = [True, True, True, True]
  rq_read_dst_req = [True, True, True, True]
  rq_read_pco_req = [True, True, True, True]

  rq_read_snu_1_req = False
  rq_read_snu_2_req = False
  rq_read_snu_3_req = False
  rq_read_snu_4_req = False

  rq_read_fwv_1_req = False
  rq_read_fwv_2_req = False
  rq_read_fwv_3_req = False
  rq_read_fwv_4_req = False

  rq_read_ver_1_req = False
  rq_read_ver_2_req = False
  rq_read_ver_3_req = False
  rq_read_ver_4_req = False

  rq_write_act_request = [False, False, False, False]
  rq_write_gto_request = [False, False, False, False]
  rq_write_atr_request = [False, False, False, False]
  rq_write_ard_request = [False, False, False, False]
  rq_write_pos_request = [False, False, False, False]
  rq_write_lbp_request = [False, False, False, False]
  rq_write_lrd_request = [False, False, False, False]
  rq_write_lbl_request = [False, False, False, False]
  rq_write_lgn_request = [False, False, False, False]
  rq_write_msc_request = [False, False, False, False]
  rq_write_mod_request = [False, False, False, False]

  rq_write_act = [-1, -1, -1, -1]
  rq_write_gto = [-1, -1, -1, -1]
  rq_write_atr = [-1, -1, -1, -1]
  rq_write_ard = [-1, -1, -1, -1]
  rq_write_for = [-1, -1, -1, -1]
  rq_write_spe = [-1, -1, -1, -1]
  rq_write_pos = [-1, -1, -1, -1]
  rq_write_lbp = [-1, -1, -1, -1]
  rq_write_lrd = [-1, -1, -1, -1]
  rq_write_lbl = [-1, -1, -1, -1]
  rq_write_lgn = [-1, -1, -1, -1]
  rq_write_msc = [-1, -1, -1, -1]
  rq_write_mod = [-1, -1, -1, -1]

  rq_write_act_previous = rq_write_act
  rq_write_gto_previous = rq_write_gto
  rq_write_atr_previous = rq_write_atr
  rq_write_ard_previous = rq_write_ard
  rq_write_for_previous = rq_write_for
  rq_write_spe_previous = rq_write_spe
  rq_write_pos_previous = rq_write_pos
  rq_write_lbp_previous = rq_write_lbp
  rq_write_lrd_previous = rq_write_lrd
  rq_write_lbl_previous = rq_write_lbl
  rq_write_lgn_previous = rq_write_lgn
  rq_write_msc_previous = rq_write_msc
  rq_write_mod_previous = rq_write_mod

  gripper_connected = [False, False, False, False]
  gripper_socket_open = [False, False, False, False]
  rq_comm_clear_socket_buffer_enabled = [True, True, True, True]
  rq_comm_check_counter = 0
  rq_gripper_communication_thread_started = False

  thread rq_gripper_communication():
      rq_comm_read_constants()
      rq_comm_read_variables()
      rq_comm_initialize_write_values()

      while(True):
          rq_comm_clear_socket_buffer()
          rq_comm_check()
          rq_comm_read_variables()
          rq_comm_write_variables()

          rq_gripper_communication_thread_started = True
          sleep(0.008)
      end
  end

  def rq_socket_to_index(gripper_socket="1"):
      # Patch in case gripper_socket is an integer
      gripper_socket_string = str_cat("", gripper_socket)

      if(gripper_socket_string == "1"):
          return 0
      elif(gripper_socket_string == "2"):
          return 1
      elif(gripper_socket_string == "3"):
          return 2
      elif(gripper_socket_string == "4"):
          return 3
      end
      return 0
  end

  def rq_index_to_socket(index=0):
      if(index == 0):
          return "1"
      elif(index == 1):
          return "2"
      elif(index == 2):
          return "3"
      elif(index == 3):
          return "4"
      end
      return "1"
  end

  def rq_comm_check():
      index = 0
      rq_comm_check_fail_counter_max = 99999

      if(rq_comm_check_counter < 50):
          rq_comm_check_counter = rq_comm_check_counter + 1
      else:
          rq_comm_check_counter = 0

          while(index <= 3):
              socket = rq_index_to_socket(index)

              if(gripper_connected[index]):
                  # Patch in case gripper_socket is an integer
                  gripper_socket_string = str_cat("", socket)

                  sid_list = rq_get_sid(socket)
                  is_gripper_in_sid_list = rq_is_gripper_in_sid_list(gripper_socket_string, sid_list)

                  if(is_gripper_in_sid_list):
                      rq_comm_check_fail_counter[index] = 0
                  else:
                      rq_comm_check_fail_counter[index] = rq_comm_check_fail_counter[index] + 1
                  end

                  if(rq_comm_check_fail_counter[index] > rq_comm_check_fail_counter_max):
                      message = str_cat("Communication lost with Robotiq's Gripper Slave ID ", gripper_socket_string)
                      popup(message, "Communication Error", False, True, True)
                  end
              end
              index = index + 1
          end
      end
  end

  def rq_init_comm_if_connected(gripper_sid=9, gripper_socket="1"):
      if(not is_gripper_socket_open(gripper_socket)):
        open_gripper_socket(gripper_socket)
      end

      socket_sid_set = rq_set_sid(gripper_sid, gripper_socket)

      if(socket_sid_set):
          # Patch in case gripper_socket is an integer
          gripper_socket_string = str_cat("", gripper_socket)

          sid_list = rq_get_sid(gripper_socket)
          is_gripper_in_sid_list = rq_is_gripper_in_sid_list(gripper_socket_string, sid_list)

          if(is_gripper_in_sid_list):
              rq_set_gripper_connected(gripper_socket_string)
              return True
          end
      end

      return False
  end

  def open_gripper_socket(gripper_socket="1"):
      is_open = socket_open(rq_gripper_socket_ip_address, rq_gripper_socket_port, gripper_socket)
      set_gripper_socket_open(gripper_socket, is_open)
  end

  def rq_close_gripper_socket(gripper_socket="1"):
      socket_close(gripper_socket)
      set_gripper_socket_open(gripper_socket, False)
      rq_set_gripper_connected(gripper_socket, False)
  end


  def is_gripper_socket_open(gripper_socket="1"):
      return gripper_socket_open[rq_socket_to_index(gripper_socket)]
  end

  def set_gripper_socket_open(gripper_socket, is_open):
      gripper_socket_open[rq_socket_to_index(gripper_socket)] = is_open
  end

  def rq_set_gripper_connected(gripper_socket="1", connected = True):
      gripper_connected[rq_socket_to_index(gripper_socket)] = connected
  end

  def rq_is_gripper_connected(gripper_id="1"):
      return gripper_connected[rq_socket_to_index(gripper_id)]
  end

  def rq_set_sid(gripper_sid=9, gripper_socket="1"):
      socket_set_var("SID", gripper_sid,  gripper_socket)
      ack = socket_read_byte_list(3, gripper_socket)
      return is_ack(ack)
  end

  def rq_gripper_enable_scan(enable, gripper_socket="1"):
      socket_set_var("MUTE", not enable,  gripper_socket)
      ack = socket_read_byte_list(3, gripper_socket)
      return is_ack(ack)
  end

  def rq_gripper_enable_tool(enable, gripper_socket="1"):
      socket_set_var("TOOL", enable,  gripper_socket)
      ack = socket_read_byte_list(3, gripper_socket)
      return is_ack(ack)
  end

  def rq_get_sid(gripper_socket="1"):
      socket_send_string("GET SID", gripper_socket)
      sid_list = socket_read_byte_list(17, gripper_socket)
      return sid_list
  end

  def rq_wait_for_gripper_connected():
      gripper_socket = "gripper_conn_socket"
      socket_open(rq_gripper_socket_ip_address, rq_gripper_socket_port, gripper_socket)

      remainingRetries = 2000
      sid_list = rq_get_sid(gripper_socket)
      gripper_is_connected = rq_is_any_gripper_connected(sid_list)

      while(not gripper_is_connected and remainingRetries > 0):
          remainingRetries = remainingRetries - 1
          sid_list = rq_get_sid(gripper_socket)
          gripper_is_connected = rq_is_any_gripper_connected(sid_list)
      end

      socket_close(gripper_socket)
  end

  def rq_is_any_gripper_connected(sid_list):
      is_gripper_1_connected = rq_is_gripper1_in_sid_list(sid_list)
      is_gripper_2_connected = rq_is_gripper2_in_sid_list(sid_list)
      is_gripper_3_connected = rq_is_gripper3_in_sid_list(sid_list)
      is_gripper_4_connected = rq_is_gripper4_in_sid_list(sid_list)

      return is_gripper_1_connected or is_gripper_2_connected or is_gripper_3_connected or is_gripper_4_connected
  end

  def rq_is_gripper_ascii_in_sid_list(gripper_ascii_sid, sid_list):
      sid_list_length = sid_list[0]
      sid_list_empty_length = 2

      if (sid_list_length <= sid_list_empty_length):
          return False
      end

      sid1 = sid_list[2]
      sid2 = sid_list[5]
      sid3 = sid_list[8]
      sid4 = sid_list[11]

      return sid1 == gripper_ascii_sid or sid2 == gripper_ascii_sid or sid3 == gripper_ascii_sid or sid4 == gripper_ascii_sid
  end

  def rq_is_gripper_in_sid_list(gripper_socket_string, sid_list):
      if(gripper_socket_string == "1"):
          return rq_is_gripper1_in_sid_list(sid_list)
      elif(gripper_socket_string == "2"):
          return rq_is_gripper2_in_sid_list(sid_list)
      elif(gripper_socket_string == "3"):
          return rq_is_gripper3_in_sid_list(sid_list)
      elif(gripper_socket_string == "4"):
          return rq_is_gripper4_in_sid_list(sid_list)
      end
      return False
  end

  def rq_is_gripper1_in_sid_list(sid_list):
      gripper_1_sid_ascii = 57
      return rq_is_gripper_ascii_in_sid_list(gripper_1_sid_ascii, sid_list)
  end

  def rq_is_gripper2_in_sid_list(sid_list):
      gripper_2_sid_ascii = 50
      return rq_is_gripper_ascii_in_sid_list(gripper_2_sid_ascii, sid_list)
  end

  def rq_is_gripper3_in_sid_list(sid_list):
      gripper_3_sid_ascii = 51
      return rq_is_gripper_ascii_in_sid_list(gripper_3_sid_ascii, sid_list)
  end

  def rq_is_gripper4_in_sid_list(sid_list):
      gripper_4_sid_ascii = 52
      return rq_is_gripper_ascii_in_sid_list(gripper_4_sid_ascii, sid_list)
  end

  def rq_comm_clear_socket_buffer():
      index = 0

      while(index <= 3):
          socket = rq_index_to_socket(index)

          if(gripper_connected[index] and rq_comm_clear_socket_buffer_enabled[index]):
              byte_in_buffer = socket_read_byte_list(1, socket, 0.002)
              while(byte_in_buffer[0] >= 1):
                  byte_in_buffer = socket_read_byte_list(1, socket, 0.002)
              end
              rq_comm_clear_socket_buffer_enabled[index] = False
          end
          index = index + 1
      end
  end

  def rq_comm_initialize_write_values():
      index = 0

      while(index <= 3):
          socket = rq_index_to_socket(index)

          if(gripper_connected[index]):

              if(rq_write_act[index] == -1 and rq_read_act[index] != -1):
                  rq_write_act[index] = rq_read_act[index]
                  rq_write_act_previous[index] = rq_read_act[index]
              elif(rq_write_act_previous[index] == -1 and rq_read_act[index] != -1):
                  rq_write_act_previous[index] = rq_read_act[index]
              end

              if(rq_write_gto[index] == -1 and rq_read_gto[index] != -1):
                  rq_write_gto[index] = rq_read_gto[index]
                  rq_write_gto_previous[index] = rq_read_gto[index]
              elif(rq_write_gto_previous[index] == -1 and rq_read_gto[index] != -1):
                  rq_write_gto_previous[index] = rq_read_gto[index]
              end

              if(rq_write_for[index] == -1 and rq_read_for[index] != -1):
                  rq_write_for[index] = rq_read_for[index]
                  rq_write_for_previous[index] = rq_read_for[index]
              elif(rq_write_for_previous[index] == -1 and rq_read_for[index] != -1):
                  rq_write_for_previous[index] = rq_read_for[index]
              end

              if(rq_write_spe[index] == -1 and rq_read_spe[index] != -1):
                  rq_write_spe[index] = rq_read_spe[index]
                  rq_write_spe_previous[index] = rq_read_spe[index]
              elif(rq_write_spe_previous[index] == -1 and rq_read_spe[index] != -1):
                  rq_write_spe_previous[index] = rq_read_spe[index]
              end

              if(rq_write_pos[index] == -1 and rq_read_pos[index] != -1):
                  rq_write_pos[index] = rq_read_pos[index]
                  rq_write_pos_previous[index] = rq_read_pos[index]
              elif(rq_write_pos_previous[index] == -1 and rq_read_pos[index] != -1):
                  rq_write_pos_previous[index] = rq_read_pos[index]
              end

              if(rq_write_lbp[index] == -1 and rq_read_lbp[index] != -1):
                  rq_write_lbp[index] = rq_read_lbp[index]
                  rq_write_lbp_previous[index] = rq_read_lbp[index]
              elif(rq_write_lbp_previous[index] == -1 and rq_read_lbp[index] != -1):
                  rq_write_lbp_previous[index] = rq_read_lbp[index]
              end

              if(rq_write_lrd[index] == -1 and rq_read_lrd[index] != -1):
                  rq_write_lrd[index] = rq_read_lrd[index]
                  rq_write_lrd_previous[index] = rq_read_lrd[index]
              elif(rq_write_lrd_previous[index] == -1 and rq_read_lrd[index] != -1):
                  rq_write_lrd_previous[index] = rq_read_lrd[index]
              end

              if(rq_write_lbl[index] == -1 and rq_read_lbl[index] != -1):
                  rq_write_lbl[index] = rq_read_lbl[index]
                  rq_write_lbl_previous[index] = rq_read_lbl[index]
              elif(rq_write_lbl_previous[index] == -1 and rq_read_lbl[index] != -1):
                  rq_write_lbl_previous[index] = rq_read_lbl[index]
              end

              if(rq_write_lgn[index] == -1 and rq_read_lgn[index] != -1):
                  rq_write_lgn[index] = rq_read_lgn[index]
                  rq_write_lgn_previous[index] = rq_read_lgn[index]
              elif(rq_write_lgn_previous[index] == -1 and rq_read_lgn[index] != -1):
                  rq_write_lgn_previous[index] = rq_read_lgn[index]
              end

              if(rq_write_msc[index] == -1 and rq_read_msc[index] != -1):
                  rq_write_msc[index] = rq_read_msc[index]
                  rq_write_msc_previous[index] = rq_read_msc[index]
              elif(rq_write_msc_previous[index] == -1 and rq_read_msc[index] != -1):
                  rq_write_msc_previous[index] = rq_read_msc[index]
              end

              if(rq_write_mod[index] == -1 and rq_read_mod[index] != -1):
                  rq_write_mod[index] = rq_read_mod[index]
                  rq_write_mod_previous[index] = rq_read_mod[index]
              elif(rq_write_mod_previous[index] == -1 and rq_read_mod[index] != -1):
                  rq_write_mod_previous[index] = rq_read_mod[index]
              end

          end
          index = index + 1
      end
  end

  def rq_comm_set_var(var, value=0, gripper_socket="1"):
      socket_set_var(var, value, gripper_socket)
      return socket_read_byte_list(3, gripper_socket)
  end

  def rq_comm_set_pos_spe_for(pos=0, speed=0, force=0, gripper_socket="1"):
      socket_send_string("SET POS", gripper_socket)
      socket_send_byte(32, gripper_socket)
      socket_send_string(pos, gripper_socket)
      socket_send_byte(32, gripper_socket)
      socket_send_string("SPE", gripper_socket)
      socket_send_byte(32, gripper_socket)
      socket_send_string(speed, gripper_socket)
      socket_send_byte(32, gripper_socket)
      socket_send_string("FOR", gripper_socket)
      socket_send_byte(32, gripper_socket)
      socket_send_string(force, gripper_socket)
      socket_send_byte(10, gripper_socket)
      return socket_read_byte_list(3, gripper_socket)
  end

  def rq_comm_read_variables():
      index = 0

      while(index <= 3):
          socket = rq_index_to_socket(index)

          if(gripper_connected[index]):

              if(rq_read_act_req[index]):
                  rq_read_act[index] = socket_get_var("ACT", socket)
                  rq_read_act_req[index] = False
              end

              if(rq_read_gto_req[index]):
                  rq_read_gto[index] = socket_get_var("GTO", socket)
                  rq_read_gto_req[index] = False
              end

              if(rq_read_pre_req[index]):
                  rq_read_pre[index] = socket_get_var("PRE", socket)
                  rq_read_pre_req[index] = False
              end

              if(rq_read_pos_req[index]):
                  rq_read_pos[index] = socket_get_var("POS", socket)
                  rq_read_pos_req[index] = False
              end

              if(rq_read_spe_req[index]):
                  rq_read_spe[index] = socket_get_var("SPE", socket)
                  rq_read_spe_req[index] = False
              end

              if(rq_read_for_req[index]):
                  rq_read_for[index] = socket_get_var("FOR", socket)
                  rq_read_for_req[index] = False
              end

              if(rq_read_obj_req[index]):
                  rq_read_obj[index] = socket_get_var("OBJ", socket)
                  rq_read_obj_req[index] = False
              end

              if(rq_read_sta_req[index]):
                  rq_read_sta[index] = socket_get_var("STA", socket)
                  rq_read_sta_req[index] = False
              end

              if(rq_read_mod_req[index]):
                  rq_read_mod[index] = socket_get_var("MOD", socket)
                  rq_read_mod_req[index] = False
              end

              if(rq_read_flt_req[index]):
                  rq_read_flt[index] = socket_get_var("FLT",socket)
                  rq_read_flt_req[index] = False
              end

              if(rq_read_lbp_req[index]):
                  rq_read_lbp[index] = socket_get_var("LBP", socket)
                  rq_read_lbp_req[index] = False
              end

              if(rq_read_lrd_req[index]):
                  rq_read_lrd[index] = socket_get_var("LRD", socket)
                  rq_read_lrd_req[index] = False
              end

              if(rq_read_lbl_req[index]):
                  rq_read_lbl[index] = socket_get_var("LBL",socket)
                  rq_read_lbl_req[index] = False
              end

              if(rq_read_lgn_req[index]):
                  rq_read_lgn[index] = socket_get_var("LGN", socket)
                  rq_read_lgn_req[index] = False
              end

              if(rq_read_msc_req[index]):
                  rq_read_msc[index] = socket_get_var("MSC", socket)
                  rq_read_msc_req[index] = False
              end

              if(rq_read_cou_req[index]):
                  rq_read_cou[index] = socket_get_var("COU", socket)
                  rq_read_cou_req[index] = False
              end

              if(rq_read_ncy_req[index]):
                  rq_read_ncy[index] = socket_get_var("NCY", socket)
                  rq_read_ncy_req[index] = False
              end

              if(rq_read_dst_req[index]):
                  rq_read_dst[index] = socket_get_var("DST", socket)
                  rq_read_dst_req[index] = False
              end

              if(rq_read_pco_req[index]):
                  rq_read_pco[index] = socket_get_var("PCO", socket)
                  rq_read_pco_req[index] = False
              end
          end
          index = index + 1
      end
  end

  def rq_comm_read_constants():

      if(gripper_connected[0]):
          while(rq_read_snu_1 == rq_string_initial_value):
              socket_send_string("GET SNU", "1")
              rq_read_snu_1 = socket_read_string("1")
          end

          while(rq_read_fwv_1 == rq_string_initial_value):
              socket_send_string("GET FWV", "1")
              rq_read_fwv_1 = socket_read_string("1")
          end

          while(rq_read_ver_1 == rq_string_initial_value):
              socket_send_string("GET VER", "1")
              rq_read_ver_1 = socket_read_string("1")
          end
      end

      if(gripper_connected[1]):
          while(rq_read_snu_2 == rq_string_initial_value):
              socket_send_string("GET SNU", "2")
              rq_read_snu_2 = socket_read_string("2")
          end

          while(rq_read_fwv_2 == rq_string_initial_value):
              socket_send_string("GET FWV", "2")
              rq_read_fwv_2 = socket_read_string("2")
          end

          while(rq_read_ver_2 == rq_string_initial_value):
              socket_send_string("GET VER", "2")
              rq_read_ver_2 = socket_read_string("2")
          end
      end

      if(gripper_connected[2]):
          while(rq_read_snu_3 == rq_string_initial_value):
              socket_send_string("GET SNU", "3")
              rq_read_snu_3 = socket_read_string("3")
          end

          while(rq_read_fwv_3 == rq_string_initial_value):
              socket_send_string("GET FWV", "3")
              rq_read_fwv_3 = socket_read_string("3")
          end

          while(rq_read_ver_3 == rq_string_initial_value):
              socket_send_string("GET VER", "3")
              rq_read_ver_3 = socket_read_string("3")
          end
      end

      if(gripper_connected[3]):
          while(rq_read_snu_4 == rq_string_initial_value):
              socket_send_string("GET SNU", "4")
              rq_read_snu_4 = socket_read_string("4")
          end

          while(rq_read_fwv_4 == rq_string_initial_value):
              socket_send_string("GET FWV", "4")
              rq_read_fwv_4 = socket_read_string("4")
          end

          while(rq_read_ver_4 == rq_string_initial_value):
              socket_send_string("GET VER", "4")
              rq_read_ver_4 = socket_read_string("4")
          end
      end
  end

  def rq_comm_write_variables():
      index = 0

      while(index <= 3):
          socket = rq_index_to_socket(index)

          if(gripper_connected[index]):

              if(rq_write_act_request[index]):
                  if(is_ack(rq_comm_set_var("ACT", rq_write_act[index], socket))):
                      rq_write_act_previous[index] = rq_write_act[index]
                      rq_write_act_request[index] = False
                  end
              end

              if(rq_write_gto_request[index]):
                  if(is_ack(rq_comm_set_var("GTO", rq_write_gto[index], socket))):
                      rq_write_gto_previous[index] = rq_write_gto[index]
                      rq_write_gto_request[index] = False
                  end
              end

              if(rq_write_atr_request[index]):
                  if(is_ack(rq_comm_set_var("ATR", rq_write_atr[index], socket))):
                      rq_write_atr_previous[index] = rq_write_atr[index]
                      rq_write_atr_request[index] = False
                  end
              end

              if(rq_write_ard_request[index]):
                  if(is_ack(rq_comm_set_var("ARD", rq_write_ard[index], socket))):
                      rq_write_ard_previous[index] = rq_write_ard[index]
                      rq_write_ard_request[index] = False
                  end
              end

              if(rq_write_pos_request[index]):
                  if(is_ack(rq_comm_set_pos_spe_for(rq_write_pos[index], rq_write_spe[index], rq_write_for[index], socket))):
                      rq_write_pos_previous[index] = rq_write_pos[index]
                      rq_write_spe_previous[index] = rq_write_spe[index]
                      rq_write_for_previous[index] = rq_write_for[index]
                      rq_write_pos_request[index] = False
                  end
              end

              if(rq_write_lbp_request[index]):
                  if(is_ack(rq_comm_set_var("LBP", rq_write_lbp[index], socket))):
                      rq_write_lbp_previous[index] = rq_write_lbp[index]
                      rq_write_lbp_request[index] = False
                  end
              end

              if(rq_write_lrd_request[index]):
                  if(is_ack(rq_comm_set_var("LRD", rq_write_lrd[index], socket))):
                      rq_write_lrd_previous[index] = rq_write_lrd[index]
                      rq_write_lrd_request[index] = False
                  end
              end

              if(rq_write_lbl_request[index]):
                  if(is_ack(rq_comm_set_var("LBL", rq_write_lbl[index], socket))):
                      rq_write_lbl_previous[index] = rq_write_lbl[index]
                      rq_write_lbl_request[index] = False
                  end
              end

              if(rq_write_lgn_request[index]):
                  if(is_ack(rq_comm_set_var("LGN", rq_write_lgn[index], socket))):
                      rq_write_lgn_previous[index] = rq_write_lgn[index]
                      rq_write_lgn_request[index] = False
                  end
              end

              if(rq_write_msc_request[index]):
                  if(is_ack(rq_comm_set_var("MSC", rq_write_msc[index], socket))):
                      rq_write_msc_previous[index] = rq_write_msc[index]
                      rq_write_msc_request[index] = False
                  end
              end

              if(rq_write_mod_request[index]):
                  if(is_ack(rq_comm_set_var("MOD", rq_write_mod[index], socket))):
                      rq_write_mod_previous[index] = rq_write_mod[index]
                      rq_write_mod_request[index] = False
                  end
              end
          end
          index = index + 1
      end
  end

  def rq_activate(gripper_socket="1"):
      if (not rq_is_gripper_activated(gripper_socket)):
          rq_reset(gripper_socket)

          while(not rq_get_var("ACT", 1, gripper_socket) == 0 or not rq_get_var("STA", 1, gripper_socket) == 0):
              rq_reset(gripper_socket)
              sleep(0.008)
          end

          rq_set_var("ACT",1, gripper_socket)
      end
  end

  def rq_activate_and_wait(gripper_socket="1"):
      if (not rq_is_gripper_activated(gripper_socket)):
          rq_activate(gripper_socket)
          sleep(1.0)

          while(not rq_get_var("ACT", 1, gripper_socket) == 1 or not rq_get_var("STA", 1, gripper_socket) == 3):
              sleep(0.1)
          end

          sleep(0.5)
      end
  end

  def rq_activate_all_grippers(reset=False):
      if(gripper_connected[0]):
          rq_reset_and_activate("1", reset)
      end

      if(gripper_connected[1]):
          rq_reset_and_activate("2", reset)
      end

      if(gripper_connected[2]):
          rq_reset_and_activate("3", reset)
      end

      if(gripper_connected[3]):
          rq_reset_and_activate("4", reset)
      end
  end

  def rq_reset_and_activate(gripper_socket="1", reset=False):
      if(reset):
          rq_reset(gripper_socket)
          rq_activate_and_wait(gripper_socket)
      elif(not rq_is_gripper_activated(gripper_socket)):
          rq_activate_and_wait(gripper_socket)
      end
  end

  def rq_reset(gripper_socket="1"):
      rq_set_var("ACT", 0, gripper_socket)
      rq_set_var("ATR", 0, gripper_socket)

      while(not rq_get_var("ACT", 1, gripper_socket) == 0 or not rq_get_var("STA", 1, gripper_socket) == 0):
          rq_set_var("ACT", 0, gripper_socket)
          rq_set_var("ATR", 0, gripper_socket)
          sleep(0.008)
      end

      sleep(0.5)
  end

  def rq_auto_release_open_and_wait(gripper_socket="1"):
      rq_set_var("ATR",0, gripper_socket)
      rq_set_var("ARD",0, gripper_socket)
      rq_set_var("ACT",1, gripper_socket)
      sleep(0.1)
      rq_set_var("ATR",1, gripper_socket)

      rq_wait_autorelease_completed(gripper_socket)
  end

  def rq_auto_release_close_and_wait(gripper_socket="1"):
      rq_set_var("ATR",0, gripper_socket)
      rq_set_var("ARD",1, gripper_socket)
      rq_set_var("ACT",1, gripper_socket)
      sleep(0.1)
      rq_set_var("ATR",1, gripper_socket)

      rq_wait_autorelease_completed(gripper_socket)
  end

  def rq_wait_autorelease_completed(gripper_socket="1"):
      remainingRetries = 20
      gFLT = rq_get_var("FLT", 2, gripper_socket)

      while(not is_FLT_autorelease_in_progress(gFLT) and remainingRetries > 0):
          remainingRetries = remainingRetries - 1
          gFLT = rq_get_var("FLT", 2, gripper_socket)
          sleep(0.1)
      end

      remainingRetries = 100
      gFLT = rq_get_var("FLT", 2, gripper_socket)

      while(not is_FLT_autorelease_completed(gFLT) and remainingRetries > 0):
          remainingRetries = remainingRetries - 1
          gFLT = rq_get_var("FLT", 2, gripper_socket)
          sleep(0.1)
      end
  end

  def rq_set_force(force, gripper_socket="1"):
      local force = floor(scale(force, [0, 255], [0.0, 255.0]))
      rq_set_var("FOR", force, gripper_socket)
  end

  def rq_set_speed(speed, gripper_socket="1"):
      local speed = floor(scale(speed, [0, 255], [0.0, 255.0]))
      rq_set_var("SPE", speed, gripper_socket)
  end

  def rq_open(gripper_socket="1"):
      rq_move(0, gripper_socket)
  end

  def rq_close(gripper_socket="1"):
      rq_move(255, gripper_socket)
  end

  def rq_open_and_wait(gripper_socket="1"):
      rq_move_and_wait(0, gripper_socket)
  end

  def rq_close_and_wait(gripper_socket="1"):
      rq_move_and_wait(255, gripper_socket)
  end

  def rq_move(pos, gripper_socket="1"):
      rq_set_pos(pos, gripper_socket)
      rq_go_to(gripper_socket)
  end

  def rq_move_and_wait(pos, gripper_socket="1"):
      rq_move(pos, gripper_socket)

      while (not rq_is_motion_complete(gripper_socket)):
          # wait for motion completed
          sleep(0.008)
      end
  end

  def rq_wait_for_pos_request(pos, gripper_socket="1"):
      gPRE = rq_get_var("PRE", 3, gripper_socket)

      while (gPRE != pos):
          rq_set_var("POS", pos, gripper_socket)
          sleep(0.008)
          gPRE = rq_get_var("PRE", 3, gripper_socket)
      end
  end

  def rq_wait_pos_spe_for_request(pos, speed, force, gripper_socket="1"):
      gPRE = rq_get_var("PRE", 3, gripper_socket)

      while (gPRE != pos):
          rq_set_pos_spe_for_var(pos, speed, force, gripper_socket)
          sleep(0.008)
          gPRE = rq_get_var("PRE", 3, gripper_socket)
      end
  end

  def rq_wait_for_pos(pos, gripper_socket="1"):
      rq_wait_for_pos_request(pos, gripper_socket)

      # Wait for the gripper motion to complete
      while (not rq_is_motion_complete(gripper_socket)):
          # wait for motion completed
          sleep(0.008)
          rq_set_var("GTO", 1, gripper_socket)
      end
  end

  def rq_wait(gripper_socket="1"):
      # Wait for the gripper motion to complete
      while (not rq_is_motion_complete(gripper_socket)):
          sleep(0.008)
          # The following patch is for Robotiq's Camera issue when communication is lost, but not the activation
          # the communication driver reset the GTO bit
          rq_set_var("GTO", 1, gripper_socket)
      end
  end

  def rq_wait_for_object_detected(gripper_socket="1"):
      # Wait the object detection
      while (not rq_is_object_detected(gripper_socket)):
          sleep(0.008)
      end
  end

  # set the position
  def rq_set_pos(pos, gripper_socket="1"):
      local pos = floor(scale(pos, [0, 255], [0.0, 255.0]))
      rq_set_var("POS", pos, gripper_socket)
      rq_wait_for_pos_request(pos, gripper_socket)
  end

  def rq_set_pos_spd_for(pos, speed, force, gripper_socket="1"):
      local pos = floor(scale(pos, [0, 255], [0.0, 255.0]))
      local speed = floor(scale(speed, [0, 255], [0.0, 255.0]))
      local force = floor(scale(force, [0, 255], [0.0, 255.0]))

      rq_set_pos_spe_for_var(pos, speed, force, gripper_socket)
      rq_wait_pos_spe_for_request(pos, speed, force, gripper_socket)
  end

  def rq_set_gripper_max_current_mA(current_mA, gripper_socket="1"):
      current = floor(current_mA / 10)

      rq_set_var("MSC", current, gripper_socket)
      current_read = rq_get_var("MSC", 1, gripper_socket)

      while(current_read != current):
          rq_set_var("MSC", current, gripper_socket)
          current_read = rq_get_var("MSC", 1, gripper_socket)
      end
  end

  def rq_set_gripper_mode(mode, gripper_socket="1"):
      rq_set_var("MOD", mode, gripper_socket)
  end

  def rq_set_gripper_max_cur(current_mA, gripper_socket="1"):
      rq_set_gripper_max_current_mA(current_mA, gripper_socket)
  end

  def rq_get_gripper_max_current_mA(gripper_socket="1"):
      current = rq_get_var("MSC", 1, gripper_socket)

      if(current == -1):
          current_mA = current
      else:
          current_mA = current * 10
      end

      return current_mA
  end

  def rq_get_gripper_max_cur(gripper_socket="1"):
      return rq_get_gripper_max_current_mA(gripper_socket)
  end

  def rq_set_max_current_for_all_grippers():
      current_mA = rq_get_max_current_mA()

      if(gripper_connected[0]):
          rq_set_gripper_max_current_mA(current_mA, "1")
      end

      if(gripper_connected[1]):
          rq_set_gripper_max_current_mA(current_mA, "2")
      end

      if(gripper_connected[2]):
          rq_set_gripper_max_current_mA(current_mA, "3")
      end

      if(gripper_connected[3]):
          rq_set_gripper_max_current_mA(current_mA, "4")
      end
  end

  def rq_get_max_current_mA():
      max_current_mA = 0

      if(rq_current_limit_enabled):
          nb_connected_grippers = rq_get_nb_connected_grippers()

          if(nb_connected_grippers == 1):
              max_current_mA = 600
          elif(nb_connected_grippers > 1):
              max_current_mA = 450
          end
      else:

      end

      return max_current_mA
  end

  def rq_get_nb_connected_grippers():
      nb_connected_grippers = 0

      if(gripper_connected[0]):
          nb_connected_grippers = nb_connected_grippers + 1
      end

      if(gripper_connected[1]):
          nb_connected_grippers = nb_connected_grippers + 1
      end

      if(gripper_connected[2]):
          nb_connected_grippers = nb_connected_grippers + 1
      end

      if(gripper_connected[3]):
          nb_connected_grippers = nb_connected_grippers + 1
      end

      return nb_connected_grippers
  end

  def rq_list_of_bytes_to_value(list_of_bytes):
      value = -1

      # response list length
      if (list_of_bytes[0] == 1):
          value = list_of_bytes[1] - 48
      elif (list_of_bytes[0] == 2):
          value = (list_of_bytes[1] - 48) * 10 + (list_of_bytes[2] - 48)
      elif (list_of_bytes[0] == 3):
          value = (list_of_bytes[1] - 48) * 100 + (list_of_bytes[2] - 48) * 10 + (list_of_bytes[3] - 48)
      end

      return value
  end

  def rq_is_motion_complete(gripper_socket="1"):
      gOBJ = rq_get_var("OBJ", 1, gripper_socket)
      sleep(0.008)
      return is_OBJ_gripper_at_position(gOBJ) or is_OBJ_object_detected(gOBJ)
  end

  def rq_is_gripper_activated(gripper_socket="1"):
      gSTA = rq_get_var("STA", 1, gripper_socket)
      sleep(0.008)
      return is_STA_gripper_activated(gSTA)
  end

  def rq_is_object_detected(gripper_socket="1"):
      gOBJ = rq_get_var("OBJ", 1, gripper_socket)
      sleep(0.008)
      return is_OBJ_object_detected(gOBJ)
  end

  def rq_current_pos(gripper_socket="1"):
      gPOS = rq_get_var("POS", 1, gripper_socket)
      sleep(0.008)
      return gPOS
  end

  def rq_motor_current(gripper_socket="1"):
      rq_current = rq_get_var("COU", 1, gripper_socket)
      sleep(0.008)
      return rq_current * 10
  end

  def rq_print_connected_grippers():
      if(gripper_connected[0]):
          textmsg("Gripper 1 : ", "connected and socket open.")
      end

      if (gripper_connected[1]):
          textmsg("Gripper 2 : ", "connected and socket open.")
      end

      if (gripper_connected[2]):
          textmsg("Gripper 3 : ", "connected and socket open.")
      end

      if (gripper_connected[3]):
          textmsg("Gripper 4 : ", "connected and socket open.")
      end
  end

  def rq_print_gripper_fault_code(gripper_socket="1"):
      gFLT = rq_get_var("FLT", 2, gripper_socket)

      if(is_FLT_no_fault(gFLT)):
          textmsg("Gripper Fault : ", "No Fault (0x00)")
      elif (is_FLT_action_delayed(gFLT)):
          textmsg("Gripper Fault : ", "Priority Fault: Action delayed, initialization must be completed prior to performing the action (0x05)")
      elif (is_FLT_not_activated(gFLT)):
          textmsg("Gripper Fault : ", "Priority Fault: The activation bit must be set prior to performing the action (0x07)")
      elif (is_FLT_over_temperature(gFLT)):
          textmsg("Gripper Fault : ", "Minor Fault: Maximum operating temperature exceeded (≥ 85°C internally), let cool down (below 80°C) (0x08)")
      elif (is_FLT_no_communication(gFLT)):
          textmsg("Gripper Fault : ", "Minor Fault: No communication during at least 1 second (0x09)")
      elif (is_FLT_under_voltage(gFLT)):
          textmsg("Gripper Fault : ", "Major Fault: Under minimum operating voltage (0x0A)")
      elif (is_FLT_autorelease_in_progress(gFLT)):
          textmsg("Gripper Fault : ", "Major Fault: Automatic release in progress (0x0B)")
      elif (is_FLT_internal_fault(gFLT)):
          textmsg("Gripper Fault : ", "Major Fault: Internal fault; contact support@robotiq.com (0x0C)")
      elif (is_FLT_activation_error(gFLT)):
          textmsg("Gripper Fault : ", "Major Fault: Activation fault; verify that no interference or other error occurred (0x0D)")
      elif (is_FLT_overcurrent(gFLT)):
          textmsg("Gripper Fault : ", "Major Fault: Overcurrent triggered (0x0E)")
      elif (is_FLT_autorelease_completed(gFLT)):
          textmsg("Gripper Fault : ", "Major Fault: Automatic release completed (0x0F)")
      else:
          textmsg("Gripper Fault : ", "Unknown Fault")
      end
  end

  def rq_print_gripper_num_cycles(gripper_socket="1"):
      num_cycles = rq_get_var("NCY", 1, gripper_socket)

      if(num_cycles == -1):
          textmsg("Gripper Cycle Number : ", "Number of cycles is unreachable.")
      else:
          textmsg("Gripper Cycle Number : ", num_cycles)
      end
  end

  def rq_print_gripper_driver_state(gripper_socket="1"):
      driver_state = rq_get_var("DST", 1, gripper_socket)

      if(driver_state == 0):
          textmsg("Gripper Driver State : ", "RQ_STATE_INIT")
      elif(driver_state == 1):
          textmsg("Gripper Driver State : ", "RQ_STATE_LISTEN")
      elif(driver_state == 2):
          textmsg("Gripper Driver State : ", "RQ_STATE_READ_INFO")
      elif(driver_state == 3):
          textmsg("Gripper Driver State : ", "RQ_STATE_ACTIVATION")
      else:
          textmsg("Gripper Driver State : ", "RQ_STATE_RUN")
      end
  end

  def rq_print_gripper_serial_number(gripper_socket="1"):
      serial_number = rq_get_var_string("SNU", 1, gripper_socket)
      textmsg("Gripper Serial Number : ", serial_number)
  end

  def rq_print_gripper_firmware_version(gripper_socket="1"):
      firmware_version = rq_get_var_string("FWV", 1, gripper_socket)
      textmsg("Gripper Firmware Version : ", firmware_version)
  end

  def rq_print_gripper_driver_version(gripper_socket="1"):
      driver_version = rq_get_var_string("VER", 1, gripper_socket)
      textmsg("Gripper Driver Version : ", driver_version)
  end

  def rq_print_gripper_connection_state(gripper_socket="1"):
      connection_state = rq_get_var("PCO", 1, gripper_socket)

      if (connection_state == 0):
          textmsg("Gripper Connection State : ", "No connection problem detected")
      else:
          textmsg("Gripper Connection State : ", "Connection problem detected")
      end
  end

  # Returns True if list_of_bytes is [3, 'a', 'c', 'k']
  def is_ack(list_of_bytes):

      # list length is not 3
      if (list_of_bytes[0] != 3):
          return False
      end

      # first byte not is 'a'?
      if (list_of_bytes[1] != 97):
          return False
      end

      # first byte not is 'c'?
      if (list_of_bytes[2] != 99):
          return False
      end

      # first byte not is 'k'?
      if (list_of_bytes[3] != 107):
          return False
      end

      return True
  end

  # Returns True if list_of_bytes is not [3, 'a', 'c', 'k']
  def is_not_ack(list_of_bytes):
      if (is_ack(list_of_bytes)):
          return False
      else:
          return True
      end
  end

  def is_STA_gripper_activated (gSTA):
      if (gSTA == 3):
          return True
      end

      return False
  end

  def is_OBJ_object_detected (gOBJ):
      if (gOBJ == 1 or gOBJ == 2):
          return True
      end

      return False
  end

  def is_OBJ_gripper_at_position (gOBJ):
      if (gOBJ == 3):
          return True
      end

      return False
  end

  def is_not_OBJ_gripper_at_position (gOBJ):
      if (is_OBJ_gripper_at_position(gOBJ)):
          return False
      else:
          return True
      end
  end

  #### GTO Section ####
  def rq_stop(gripper_socket="1"):
      rq_set_var("GTO", 0, gripper_socket)
  end

  def rq_set_GTO_and_wait(value, gripper_socket="1"):
      rq_set_var("GTO" ,value, gripper_socket)
      while(not is_GTO(value, rq_get_var("GTO", 1, gripper_socket))):
        sleep(0.008)
      end
  end

  def rq_go_to(gripper_socket="1"):
      rq_set_var("GTO", 1, gripper_socket)
  end


  def is_GTO(goto_value, rGTO):
      return rGTO == goto_value
  end
  #### GTO Section ####

  def is_FLT_no_fault(gFLT):
      return gFLT == 0
  end

  def is_FLT_warning(gFLT):
      return gFLT >= 1 and gFLT <= 7
  end

  def is_FLT_faulted(gFLT):
      return gFLT >= 8
  end

  def is_FLT_action_delayed(gFLT):
      return gFLT == 5
  end

  def is_FLT_not_activated(gFLT):
      return gFLT == 7
  end

  def is_FLT_over_temperature(gFLT):
      return gFLT == 8
  end

  def is_FLT_no_communication(gFLT):
      return gFLT == 9
  end

  def is_FLT_under_voltage(gFLT):
      return gFLT == 10
  end

  def is_FLT_autorelease_in_progress(gFLT):
      return gFLT == 11
  end

  def is_FLT_internal_fault(gFLT):
      return gFLT == 12
  end

  def is_FLT_activation_error(gFLT):
      return gFLT == 13
  end

  def is_FLT_overcurrent(gFLT):
      return gFLT == 14
  end

  def is_FLT_autorelease_completed(gFLT):
      return gFLT == 15
  end

  def rq_set_var(var_name, var_value, gripper_socket="1"):
      index = rq_socket_to_index(gripper_socket)

      enter_critical

      if (var_name == "ACT"):
          rq_write_act[index] = var_value
          rq_write_act_request[index] = True
      elif (var_name == "GTO"):
          rq_write_gto[index] = var_value
          rq_write_gto_request[index] = True
      elif (var_name == "ATR"):
          rq_write_atr[index] = var_value
          rq_write_atr_request[index] = True
      elif (var_name == "ARD"):
          rq_write_ard[index] = var_value
          rq_write_ard_request[index] = True
      elif (var_name == "FOR"):
          rq_write_for[index] = var_value
          rq_write_pos_request[index] = True
      elif (var_name == "SPE"):
          rq_write_spe[index] = var_value
          rq_write_pos_request[index] = True
      elif (var_name == "POS"):
          rq_write_pos[index] = var_value
          rq_write_pos_request[index] = True
      elif (var_name == "LBP"):
          rq_write_lbp[index] = var_value
          rq_write_lbp_request[index] = True
      elif (var_name == "LRD"):
          rq_write_lrd[index] = var_value
          rq_write_lrd_request[index] = True
      elif (var_name == "LBL"):
          rq_write_lbl[index] = var_value
          rq_write_lbl_request[index] = True
      elif (var_name == "LGN"):
          rq_write_lgn[index] = var_value
          rq_write_lgn_request[index] = True
      elif (var_name == "MSC"):
          rq_write_msc[index] = var_value
          rq_write_msc_request[index] = True
      elif (var_name == "MOD"):
          rq_write_mod[index] = var_value
          rq_write_mod_request[index] = True
      end

      exit_critical

      if (var_name == "ACT"):
          while(rq_write_act_request[index]):
              sleep(0.008)
          end
      elif (var_name == "GTO"):
          while(rq_write_gto_request[index]):
              sleep(0.008)
          end
      elif (var_name == "ATR"):
          while(rq_write_atr_request[index]):
              sleep(0.008)
          end
      elif (var_name == "ARD"):
          while(rq_write_ard_request[index]):
              sleep(0.008)
          end
      elif (var_name == "FOR"):
          while(rq_write_pos_request[index]):
              sleep(0.008)
          end
      elif (var_name == "SPE"):
          while(rq_write_pos_request[index]):
              sleep(0.008)
          end
      elif (var_name == "POS"):
          while(rq_write_pos_request[index]):
              sleep(0.008)
          end
      elif (var_name == "LBP"):
          while(rq_write_lbp_request[index]):
              sleep(0.008)
          end
      elif (var_name == "LRD"):
          while(rq_write_lrd_request[index]):
              sleep(0.008)
          end
      elif (var_name == "LBL"):
          while(rq_write_lbl_request[index]):
              sleep(0.008)
          end
      elif (var_name == "LGN"):
          while(rq_write_lgn_request[index]):
              sleep(0.008)
          end
      elif (var_name == "MSC"):
          while(rq_write_msc_request[index]):
              sleep(0.008)
          end
      elif (var_name == "MOD"):
          while(rq_write_mod_request[index]):
              sleep(0.008)
          end
      end
  end

  def rq_set_pos_spe_for_var(pos, speed, force, gripper_socket="1"):
      index = rq_socket_to_index(gripper_socket)

      enter_critical

      rq_write_for[index] = force
      rq_write_spe[index] = speed
      rq_write_pos[index] = pos
      rq_write_pos_request[index] = True

      exit_critical
  end

  def rq_get_var(var_name, nbr_bytes, gripper_socket="1"):
      index = rq_socket_to_index(gripper_socket)
      var_value = -1

      if (var_name == "ACT"):
          enter_critical
          rq_read_act_req[index] = True
          exit_critical
          while(rq_read_act_req[index]):
              sleep(0.008)
          end
          var_value = rq_read_act[index]

      elif (var_name == "GTO"):
          enter_critical
          rq_read_gto_req[index] = True
          exit_critical
          while(rq_read_gto_req[index]):
              sleep(0.008)
          end
          var_value = rq_read_gto[index]

      elif (var_name == "FOR"):
          enter_critical
          rq_read_for_req[index] = True
          exit_critical
          while(rq_read_for_req[index]):
              sleep(0.008)
          end
          var_value = rq_read_for[index]

      elif (var_name == "SPE"):
          enter_critical
          rq_read_spe_req[index] = True
          exit_critical
          while(rq_read_spe_req[index]):
              sleep(0.008)
          end
          var_value = rq_read_spe[index]

      elif (var_name == "OBJ"):
          enter_critical
          rq_read_obj_req[index] = True
          exit_critical
          while(rq_read_obj_req[index]):
              sleep(0.008)
          end
          var_value = rq_read_obj[index]

      elif (var_name == "STA"):
          enter_critical
          rq_read_sta_req[index] = True
          exit_critical
          while(rq_read_sta_req[index]):
              sleep(0.008)
          end
          var_value = rq_read_sta[index]

      elif (var_name == "FLT"):
          enter_critical
          rq_read_flt_req[index] = True
          exit_critical
          while(rq_read_flt_req[index]):
              sleep(0.008)
          end
          var_value = rq_read_flt[index]

      elif (var_name == "POS"):
          enter_critical
          rq_read_pos_req[index] = True
          exit_critical
          while(rq_read_pos_req[index]):
              sleep(0.008)
          end
          var_value = rq_read_pos[index]

      elif (var_name == "PRE"):
          enter_critical
          rq_read_pre_req[index] = True
          exit_critical
          while(rq_read_pre_req[index]):
              sleep(0.008)
          end
          var_value = rq_read_pre[index]

      elif (var_name == "LBP"):
          enter_critical
          rq_read_lbp_req[index] = True
          exit_critical
          while(rq_read_lbp_req[index]):
              sleep(0.008)
          end
          var_value = rq_read_lbp[index]

      elif (var_name == "LRD"):
          enter_critical
          rq_read_lrd_req[index] = True
          exit_critical
          while(rq_read_lrd_req[index]):
              sleep(0.008)
          end
          var_value = rq_read_lrd[index]

      elif (var_name == "LBL"):
          enter_critical
          rq_read_lbl_req[index] = True
          exit_critical
          while(rq_read_lbl_req[index]):
              sleep(0.008)
          end
          var_value = rq_read_lbl[index]

      elif (var_name == "LGN"):
          enter_critical
          rq_read_lgn_req[index] = True
          exit_critical
          while(rq_read_lgn_req[index]):
              sleep(0.008)
          end
          var_value = rq_read_lgn[index]

      elif (var_name == "MSC"):
          enter_critical
          rq_read_msc_req[index] = True
          exit_critical
          while(rq_read_msc_req[index]):
              sleep(0.008)
          end
          var_value = rq_read_msc[index]

      elif (var_name == "MOD"):
          enter_critical
          rq_read_mod_req[index] = True
          exit_critical
          while(rq_read_mod_req[index]):
              sleep(0.008)
          end
          var_value = rq_read_mod[index]

      elif (var_name == "NCY"):
          enter_critical
          rq_read_ncy_req[index] = True
          exit_critical
          while(rq_read_ncy_req[index]):
              sleep(0.008)
          end
          var_value = rq_read_ncy[index]

      elif (var_name == "PCO"):
          enter_critical
          rq_read_pco_req[index] = True
          exit_critical
          while(rq_read_pco_req[index]):
              sleep(0.008)
          end
          var_value = rq_read_pco[index]

      elif (var_name == "DST"):
          enter_critical
          rq_read_dst_req[index] = True
          exit_critical
          while(rq_read_dst_req[index]):
              sleep(0.008)
          end
          var_value = rq_read_dst[index]

      end

      return var_value
  end

  def rq_get_var_string(var_name, nbr_bytes, gripper_socket="1"):
      index = rq_socket_to_index(gripper_socket)
      var_value = ""

      enter_critical

      if (var_name == "SNU"):
          if(gripper_socket == "1"):
              var_value = rq_read_snu_1
          elif(gripper_socket == "2"):
              var_value = rq_read_snu_2
          elif(gripper_socket == "3"):
              var_value = rq_read_snu_3
          elif(gripper_socket == "4"):
              var_value = rq_read_snu_4
          end
      elif (var_name == "FWV"):
          if(gripper_socket == "1"):
              var_value = rq_read_fwv_1
          elif(gripper_socket == "2"):
              var_value = rq_read_fwv_2
          elif(gripper_socket == "3"):
              var_value = rq_read_fwv_3
          elif(gripper_socket == "4"):
              var_value = rq_read_fwv_4
          end
      elif (var_name == "VER"):
          if(gripper_socket == "1"):
              var_value = rq_read_ver_1
          elif(gripper_socket == "2"):
              var_value = rq_read_ver_2
          elif(gripper_socket == "3"):
              var_value = rq_read_ver_3
          elif(gripper_socket == "4"):
              var_value = rq_read_ver_4
          end
      end

      exit_critical

      return var_value
  end

  def rq_is_object_validated(gripper_selected, gripper_socket="1"):
      if(gripper_selected):
          if(rq_is_object_detected(gripper_socket)):
              return True
          else:
              return False
          end
      else:
          return True
      end
  end

  ############################################
  # normalized functions (maps 0-100 to 0-255)
  ############################################
  def rq_set_force_norm(force_norm, gripper_socket="1"):
      force_gripper = norm_to_gripper(force_norm)
      rq_set_force(force_gripper, gripper_socket)
  end

  def rq_set_speed_norm(speed_norm, gripper_socket="1"):
      speed_gripper = norm_to_gripper(speed_norm)
      rq_set_speed(speed_gripper, gripper_socket)
  end

  def rq_move_norm(pos_norm, gripper_socket="1"):
      pos_gripper = norm_to_gripper(pos_norm)
      rq_move(pos_gripper, gripper_socket)
  end

  def rq_move_and_wait_norm(pos_norm, gripper_socket="1"):
      pos_gripper = norm_to_gripper(pos_norm)
      rq_move_and_wait(pos_gripper, gripper_socket)
  end

  def rq_set_pos_norm(pos_norm, gripper_socket="1"):
      pos_gripper = norm_to_gripper(pos_norm)
      rq_set_pos(pos_gripper, gripper_socket)
  end

  def rq_current_pos_norm(gripper_socket="1"):
      pos_gripper = rq_current_pos(gripper_socket)
      pos_norm = gripper_to_norm(pos_gripper)
      return pos_norm
  end

  def gripper_to_norm(value_gripper):
      value_norm = (value_gripper / 255) * 100
      return floor(value_norm)
  end

  def norm_to_gripper(value_norm):
      value_gripper = (value_norm / 100) * 255
      return ceil(value_gripper)
  end

  def rq_get_position():
      return rq_current_pos_norm()
  end

  def rq_gripper_led_on(gripper_socket="1"):
      rq_set_var("LBP",0, gripper_socket)
  end

  def rq_gripper_led_off(gripper_socket="1"):
      rq_set_var("LBP",1, gripper_socket)
      rq_set_var("LRD",0, gripper_socket)
      rq_set_var("LBL",0, gripper_socket)
      rq_set_var("LGN",0, gripper_socket)
  end

  def rq_gripper_led_force_red(gripper_socket="1"):
      rq_set_var("LBP",1, gripper_socket)
      rq_set_var("LRD",1, gripper_socket)
      rq_set_var("LBL",0, gripper_socket)
      rq_set_var("LGN",0, gripper_socket)
  end

  def rq_gripper_led_force_blue(gripper_socket="1"):
      rq_set_var("LBP",1, gripper_socket)
      rq_set_var("LRD",0, gripper_socket)
      rq_set_var("LBL",1, gripper_socket)
      rq_set_var("LGN",0, gripper_socket)
  end

  def rq_gripper_led_force_green(gripper_socket="1"):
      rq_set_var("LBP",1, gripper_socket)
      rq_set_var("LRD",0, gripper_socket)
      rq_set_var("LBL",0, gripper_socket)
      rq_set_var("LGN",1, gripper_socket)
  end

  def rq_gripper_led_force_purple(gripper_socket="1"):
      rq_set_var("LBP",1, gripper_socket)
      rq_set_var("LRD",1, gripper_socket)
      rq_set_var("LBL",1, gripper_socket)
      rq_set_var("LGN",0, gripper_socket)
  end

  ############################################
  # mm/inches functions
  ############################################
  gripper_closed_norm = [100, 100, 100, 100]
  gripper_open_norm = [0, 0, 0, 0]
  gripper_closed_mm = [0, 0, 0, 0]
  gripper_open_mm = [50, 50, 50, 50]

  def rq_current_pos_mm(gripper_socket=1):
      pos_gripper = rq_current_pos(gripper_socket)
      pos_mm = gripper_to_mm(pos_gripper, gripper_socket)
      return round_value_2_dec(pos_mm)
  end

  def rq_current_pos_inches(gripper_socket=1):
      pos_gripper = rq_current_pos(gripper_socket)
      pos_mm = gripper_to_mm(pos_gripper, gripper_socket)
      pos_in = pos_mm / 25.4
      return round_value_2_dec(pos_in)
  end

  def rq_move_mm(pos_mm, gripper_socket=1):
      pos_gripper = mm_to_gripper(pos_mm, gripper_socket)
      rq_move(pos_gripper, gripper_socket)
  end

  def rq_move_and_wait_mm(pos_mm, gripper_socket=1):
      pos_gripper = mm_to_gripper(pos_mm, gripper_socket)
      rq_move_and_wait(pos_gripper, gripper_socket)
  end

  def rq_move_inches(pos_in, gripper_socket=1):
      pos_mm = pos_in * 25.4
      rq_move_mm(pos_mm, gripper_socket)
  end

  def rq_move_and_wait_inches(pos_in, gripper_socket=1):
      pos_mm = pos_in * 25.4
      rq_move_and_wait_mm(pos_mm, gripper_socket)
  end

  def get_closed_norm(gripper_socket):
      return gripper_closed_norm[gripper_socket - 1]
  end

  def get_open_norm(gripper_socket):
      return gripper_open_norm[gripper_socket - 1]
  end

  def get_closed_mm(gripper_socket):
      return gripper_closed_mm[gripper_socket - 1]
  end

  def get_open_mm(gripper_socket):
      return gripper_open_mm[gripper_socket - 1]
  end

  def set_closed_norm(closed_norm, gripper_socket):
      gripper_closed_norm[to_num(gripper_socket) - 1] = closed_norm
  end

  def set_open_norm(open_norm, gripper_socket):
      gripper_open_norm[to_num(gripper_socket) - 1] = open_norm
  end

  def set_closed_mm(closed_mm, gripper_socket):
      gripper_closed_mm[to_num(gripper_socket) - 1] = closed_mm
  end

  def set_open_mm(open_mm, gripper_socket):
      gripper_open_mm[to_num(gripper_socket) - 1] = open_mm
  end

